Universal Robots URScript: Fuk_Rabbit_01D.script

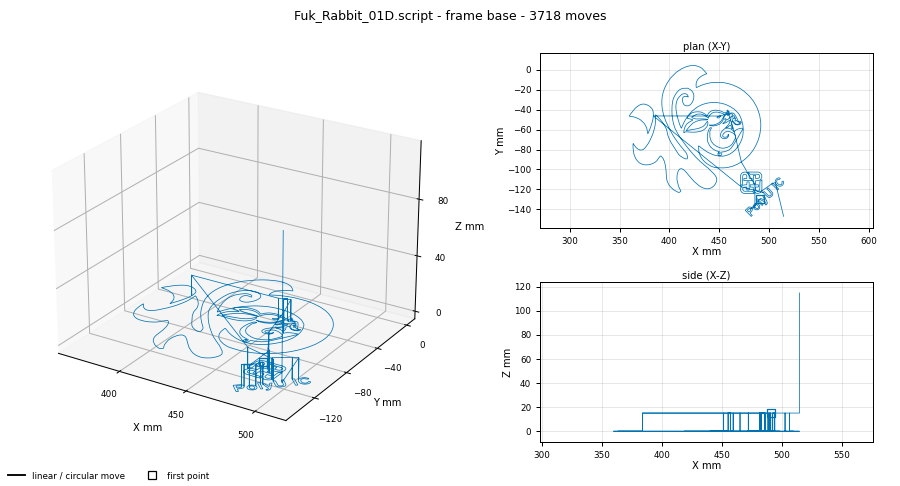
[picture p0: tool path of Fuk_Rabbit_01D.script in frame base, 3718 of 3719 moves have a stored position in this frame; points joined in program order, loops and branches not executed]
  global speed_ms    = 0.300
  global speed_rads  = 0.750
  global accel_mss   = 3.000
  global accel_radss = 1.200
  global blend_radius_m = 0.001




  # Main program:
  # Program generated by RoboDK v5.4.3 for UR10e on 11/01/2023 10:45:26
  # Using nominal kinematics.
  blend_radius_m = 0.001
  speed_ms    = 1.000
  # set_reference(p[0.514600, -0.147080, 0.000000, 0.000000, 0.000000, 1.570796])
  set_tcp(p[0.002800, -0.002800, 0.20500, 0.000000, 0.000000, 0.000000])
  movej([0.091562, -1.751682, -1.942220, -4.160080, -1.570796, -1.479235],accel_radss,speed_rads,0,0)
  movel(p[0.490670, -0.129830, 0.015000, 0.000000, -3.141593, 0.000000],accel_mss,speed_ms,0,0)

  speed_ms    = 1.000
  movel(p[0.490670, -0.129830, 0.015000, 0.000000, -3.141593, 0.000000],accel_mss,speed_ms,0,0.000)

  movel(p[0.490670, -0.129830, 0.003000, 0.000000, -3.141593, 0.000000],accel_mss,speed_ms,0,blend_radius_m)
  speed_ms    = 0.050
  movel(p[0.490670, -0.129830, -0.000100, 0.000000, -3.141593, 0.000000],accel_mss,speed_ms,0,blend_radius_m)
  speed_ms    = 0.083
  movel(p[0.491032, -0.129476, -0.000100, 0.000000, -3.141593, 0.000000],accel_mss,speed_ms,0,0.000)
  movel(p[0.491414, -0.129146, -0.000100, 0.000000, -3.141593, 0.000000],accel_mss,speed_ms,0,0.000)
  movel(p[0.491603, -0.129079, -0.000100, 0.000000, -3.141593, 0.000000],accel_mss,speed_ms,0,0.000)
  movel(p[0.491737, -0.129108, -0.000100, 0.000000, -3.141593, 0.000000],accel_mss,speed_ms,0,0.000)
  movel(p[0.492253, -0.129343, -0.000100, 0.000000, -3.141593, 0.000000],accel_mss,speed_ms,0,0.000)
  movel(p[0.492858, -0.129634, -0.000100, 0.000000, -3.141593, 0.000000],accel_mss,speed_ms,0,0.000)
  movel(p[0.493538, -0.129979, -0.000100, 0.000000, -3.141593, 0.000000],accel_mss,speed_ms,0,0.000)
  movel(p[0.494662, -0.130547, -0.000100, 0.000000, -3.141593, 0.000000],accel_mss,speed_ms,0,0.001)
  movel(p[0.495264, -0.130798, -0.000100, 0.000000, -3.141593, 0.000000],accel_mss,speed_ms,0,0.000)
  movel(p[0.495582, -0.130848, -0.000100, 0.000000, -3.141593, 0.000000],accel_mss,speed_ms,0,0.000)
  movel(p[0.495701, -0.130727, -0.000100, 0.000000, -3.141593, 0.000000],accel_mss,speed_ms,0,0.000)
  movel(p[0.495677, -0.130619, -0.000100, 0.000000, -3.141593, 0.000000],accel_mss,speed_ms,0,0.000)
  movel(p[0.495417, -0.130053, -0.000100, 0.000000, -3.141593, 0.000000],accel_mss,speed_ms,0,0.000)
  movel(p[0.495105, -0.129397, -0.000100, 0.000000, -3.141593, 0.000000],accel_mss,speed_ms,0,0.000)
  movel(p[0.494735, -0.128647, -0.000100, 0.000000, -3.141593, 0.000000],accel_mss,speed_ms,0,0.000)
  movel(p[0.494252, -0.127684, -0.000100, 0.000000, -3.141593, 0.000000],accel_mss,speed_ms,0,0.000)
  movel(p[0.493769, -0.126720, -0.000100, 0.000000, -3.141593, 0.000000],accel_mss,speed_ms,0,0.000)
  movel(p[0.494025, -0.126472, -0.000100, 0.000000, -3.141593, 0.000000],accel_mss,speed_ms,0,0.000)
  movel(p[0.494281, -0.126224, -0.000100, 0.000000, -3.141593, 0.000000],accel_mss,speed_ms,0,0.000)
  movel(p[0.494536, -0.125976, -0.000100, 0.000000, -3.141593, 0.000000],accel_mss,speed_ms,0,0.000)
  movel(p[0.494792, -0.125728, -0.000100, 0.000000, -3.141593, 0.000000],accel_mss,speed_ms,0,0.000)
  movel(p[0.495325, -0.126847, -0.000100, 0.000000, -3.141593, 0.000000],accel_mss,speed_ms,0,0.000)
  movel(p[0.495859, -0.127966, -0.000100, 0.000000, -3.141593, 0.000000],accel_mss,speed_ms,0,0.000)
  movel(p[0.496321, -0.128940, -0.000100, 0.000000, -3.141593, 0.000000],accel_mss,speed_ms,0,0.000)
  movel(p[0.496781, -0.129915, -0.000100, 0.000000, -3.141593, 0.000000],accel_mss,speed_ms,0,0.000)
  movel(p[0.497237, -0.130892, -0.000100, 0.000000, -3.141593, 0.000000],accel_mss,speed_ms,0,0.000)
  movel(p[0.497690, -0.131870, -0.000100, 0.000000, -3.141593, 0.000000],accel_mss,speed_ms,0,0.000)
  movel(p[0.498208, -0.133320, -0.000100, 0.000000, -3.141593, 0.000000],accel_mss,speed_ms,0,0.001)
  movel(p[0.498190, -0.134226, -0.000100, 0.000000, -3.141593, 0.000000],accel_mss,speed_ms,0,0.000)
  movel(p[0.497708, -0.135078, -0.000100, 0.000000, -3.141593, 0.000000],accel_mss,speed_ms,0,0.000)
  movel(p[0.497304, -0.135478, -0.000100, 0.000000, -3.141593, 0.000000],accel_mss,speed_ms,0,0.000)
  movel(p[0.497002, -0.135642, -0.000100, 0.000000, -3.141593, 0.000000],accel_mss,speed_ms,0,0.000)
  movel(p[0.496727, -0.135624, -0.000100, 0.000000, -3.141593, 0.000000],accel_mss,speed_ms,0,0.000)
  movel(p[0.496428, -0.135434, -0.000100, 0.000000, -3.141593, 0.000000],accel_mss,speed_ms,0,0.000)
  movel(p[0.496280, -0.135274, -0.000100, 0.000000, -3.141593, 0.000000],accel_mss,speed_ms,0,0.000)
  movel(p[0.496250, -0.135159, -0.000100, 0.000000, -3.141593, 0.000000],accel_mss,speed_ms,0,0.000)
  movel(p[0.496310, -0.135021, -0.000100, 0.000000, -3.141593, 0.000000],accel_mss,speed_ms,0,0.000)
  movel(p[0.496545, -0.134729, -0.000100, 0.000000, -3.141593, 0.000000],accel_mss,speed_ms,0,0.000)
  movel(p[0.496741, -0.134465, -0.000100, 0.000000, -3.141593, 0.000000],accel_mss,speed_ms,0,0.000)
  movel(p[0.496842, -0.134244, -0.000100, 0.000000, -3.141593, 0.000000],accel_mss,speed_ms,0,0.000)
  movel(p[0.496876, -0.134003, -0.000100, 0.000000, -3.141593, 0.000000],accel_mss,speed_ms,0,0.000)
  movel(p[0.496853, -0.133678, -0.000100, 0.000000, -3.141593, 0.000000],accel_mss,speed_ms,0,0.000)
  movel(p[0.496808, -0.133438, -0.000100, 0.000000, -3.141593, 0.000000],accel_mss,speed_ms,0,0.000)
  movel(p[0.496738, -0.133207, -0.000100, 0.000000, -3.141593, 0.000000],accel_mss,speed_ms,0,0.000)
  movel(p[0.496657, -0.133013, -0.000100, 0.000000, -3.141593, 0.000000],accel_mss,speed_ms,0,0.000)
  movel(p[0.496575, -0.132902, -0.000100, 0.000000, -3.141593, 0.000000],accel_mss,speed_ms,0,0.000)
  movel(p[0.496413, -0.132791, -0.000100, 0.000000, -3.141593, 0.000000],accel_mss,speed_ms,0,0.000)
  movel(p[0.495586, -0.132385, -0.000100, 0.000000, -3.141593, 0.000000],accel_mss,speed_ms,0,0.000)
  movel(p[0.494609, -0.131919, -0.000100, 0.000000, -3.141593, 0.000000],accel_mss,speed_ms,0,0.000)
  movel(p[0.493488, -0.131401, -0.000100, 0.000000, -3.141593, 0.000000],accel_mss,speed_ms,0,0.000)
  movel(p[0.492381, -0.130891, -0.000100, 0.000000, -3.141593, 0.000000],accel_mss,speed_ms,0,0.000)
  movel(p[0.491449, -0.130448, -0.000100, 0.000000, -3.141593, 0.000000],accel_mss,speed_ms,0,0.000)
  movel(p[0.490630, -0.130050, -0.000100, 0.000000, -3.141593, 0.000000],accel_mss,speed_ms,0,0.000)
  movel(p[0.490670, -0.129830, -0.000100, 0.000000, -3.141593, 0.000000],accel_mss,speed_ms,0,0.000)
  speed_ms    = 0.050
  movel(p[0.490670, -0.129830, 0.003000, 0.000000, -3.141593, 0.000000],accel_mss,speed_ms,0,blend_radius_m)
  speed_ms    = 1.000
  movel(p[0.490670, -0.129830, 0.015000, 0.000000, -3.141593, 0.000000],accel_mss,speed_ms,0,blend_radius_m)

  movel(p[0.489450, -0.130704, 0.015000, 0.000000, -3.141593, 0.000000],accel_mss,speed_ms,0,0.001)

  movel(p[0.489450, -0.130704, 0.003000, 0.000000, -3.141593, 0.000000],accel_mss,speed_ms,0,blend_radius_m)
  speed_ms    = 0.050
  movel(p[0.489450, -0.130704, -0.000100, 0.000000, -3.141593, 0.000000],accel_mss,speed_ms,0,blend_radius_m)
  speed_ms    = 0.083
  movel(p[0.490933, -0.132187, -0.000100, 0.000000, -3.141593, 0.000000],accel_mss,speed_ms,0,0.001)
  movel(p[0.492071, -0.133333, -0.000100, 0.000000, -3.141593, 0.000000],accel_mss,speed_ms,0,0.001)
  movel(p[0.493029, -0.134322, -0.000100, 0.000000, -3.141593, 0.000000],accel_mss,speed_ms,0,0.001)
  movel(p[0.493862, -0.135197, -0.000100, 0.000000, -3.141593, 0.000000],accel_mss,speed_ms,0,0.000)
  movel(p[0.493901, -0.135293, -0.000100, 0.000000, -3.141593, 0.000000],accel_mss,speed_ms,0,0.000)
  movel(p[0.493835, -0.135480, -0.000100, 0.000000, -3.141593, 0.000000],accel_mss,speed_ms,0,0.000)
  movel(p[0.493567, -0.135785, -0.000100, 0.000000, -3.141593, 0.000000],accel_mss,speed_ms,0,0.000)
  movel(p[0.493270, -0.136063, -0.000100, 0.000000, -3.141593, 0.000000],accel_mss,speed_ms,0,0.000)
  movel(p[0.493088, -0.136129, -0.000100, 0.000000, -3.141593, 0.000000],accel_mss,speed_ms,0,0.000)
  movel(p[0.492980, -0.136086, -0.000100, 0.000000, -3.141593, 0.000000],accel_mss,speed_ms,0,0.000)
  movel(p[0.492106, -0.135260, -0.000100, 0.000000, -3.141593, 0.000000],accel_mss,speed_ms,0,0.000)
  movel(p[0.491114, -0.134305, -0.000100, 0.000000, -3.141593, 0.000000],accel_mss,speed_ms,0,0.001)
  movel(p[0.489967, -0.133171, -0.000100, 0.000000, -3.141593, 0.000000],accel_mss,speed_ms,0,0.001)
  movel(p[0.488487, -0.131692, -0.000100, 0.000000, -3.141593, 0.000000],accel_mss,speed_ms,0,0.001)
  movel(p[0.487006, -0.130212, -0.000100, 0.000000, -3.141593, 0.000000],accel_mss,speed_ms,0,0.001)
  movel(p[0.487246, -0.129965, -0.000100, 0.000000, -3.141593, 0.000000],accel_mss,speed_ms,0,0.000)
  movel(p[0.487486, -0.129717, -0.000100, 0.000000, -3.141593, 0.000000],accel_mss,speed_ms,0,0.000)
  movel(p[0.487726, -0.129470, -0.000100, 0.000000, -3.141593, 0.000000],accel_mss,speed_ms,0,0.000)
  movel(p[0.487966, -0.129222, -0.000100, 0.000000, -3.141593, 0.000000],accel_mss,speed_ms,0,0.000)
  movel(p[0.489450, -0.130704, -0.000100, 0.000000, -3.141593, 0.000000],accel_mss,speed_ms,0,0.001)
  speed_ms    = 0.050
  movel(p[0.489450, -0.130704, 0.003000, 0.000000, -3.141593, 0.000000],accel_mss,speed_ms,0,blend_radius_m)
  speed_ms    = 1.000
  movel(p[0.489450, -0.130704, 0.015000, 0.000000, -3.141593, 0.000000],accel_mss,speed_ms,0,blend_radius_m)

  movel(p[0.488402, -0.134348, 0.015000, 0.000000, -3.141593, 0.000000],accel_mss,speed_ms,0,blend_radius_m)

  movel(p[0.488402, -0.134348, 0.003000, 0.000000, -3.141593, 0.000000],accel_mss,speed_ms,0,blend_radius_m)
  speed_ms    = 0.050
  movel(p[0.488402, -0.134348, -0.000100, 0.000000, -3.141593, 0.000000],accel_mss,speed_ms,0,blend_radius_m)
  speed_ms    = 0.083
  movel(p[0.489131, -0.134715, -0.000100, 0.000000, -3.141593, 0.000000],accel_mss,speed_ms,0,0.000)
  movel(p[0.489694, -0.135212, -0.000100, 0.000000, -3.141593, 0.000000],accel_mss,speed_ms,0,0.000)
  movel(p[0.490184, -0.135859, -0.000100, 0.000000, -3.141593, 0.000000],accel_mss,speed_ms,0,0.000)
  movel(p[0.490543, -0.136563, -0.000100, 0.000000, -3.141593, 0.000000],accel_mss,speed_ms,0,0.000)
  movel(p[0.490711, -0.137230, -0.000100, 0.000000, -3.141593, 0.000000],accel_mss,speed_ms,0,0.000)
  movel(p[0.490469, -0.138750, -0.000100, 0.000000, -3.141593, 0.000000],accel_mss,speed_ms,0,0.001)
  movel(p[0.489477, -0.139984, -0.000100, 0.000000, -3.141593, 0.000000],accel_mss,speed_ms,0,0.001)
  movel(p[0.488016, -0.140593, -0.000100, 0.000000, -3.141593, 0.000000],accel_mss,speed_ms,0,0.001)
  movel(p[0.486490, -0.140400, -0.000100, 0.000000, -3.141593, 0.000000],accel_mss,speed_ms,0,0.001)
  movel(p[0.485962, -0.140097, -0.000100, 0.000000, -3.141593, 0.000000],accel_mss,speed_ms,0,0.000)
  movel(p[0.485374, -0.139591, -0.000100, 0.000000, -3.141593, 0.000000],accel_mss,speed_ms,0,0.000)
  movel(p[0.484851, -0.139015, -0.000100, 0.000000, -3.141593, 0.000000],accel_mss,speed_ms,0,0.000)
  movel(p[0.484531, -0.138492, -0.000100, 0.000000, -3.141593, 0.000000],accel_mss,speed_ms,0,0.000)
  movel(p[0.484440, -0.138227, -0.000100, 0.000000, -3.141593, 0.000000],accel_mss,speed_ms,0,0.000)
  movel(p[0.484378, -0.137886, -0.000100, 0.000000, -3.141593, 0.000000],accel_mss,speed_ms,0,0.000)
  movel(p[0.484347, -0.137493, -0.000100, 0.000000, -3.141593, 0.000000],accel_mss,speed_ms,0,0.000)
  movel(p[0.484349, -0.137070, -0.000100, 0.000000, -3.141593, 0.000000],accel_mss,speed_ms,0,0.000)
  movel(p[0.484479, -0.136262, -0.000100, 0.000000, -3.141593, 0.000000],accel_mss,speed_ms,0,0.000)
  movel(p[0.484789, -0.135564, -0.000100, 0.000000, -3.141593, 0.000000],accel_mss,speed_ms,0,0.000)
  movel(p[0.485282, -0.134982, -0.000100, 0.000000, -3.141593, 0.000000],accel_mss,speed_ms,0,0.000)
  movel(p[0.485951, -0.134516, -0.000100, 0.000000, -3.141593, 0.000000],accel_mss,speed_ms,0,0.000)
  movel(p[0.486717, -0.134242, -0.000100, 0.000000, -3.141593, 0.000000],accel_mss,speed_ms,0,0.000)
  movel(p[0.487565, -0.134186, -0.000100, 0.000000, -3.141593, 0.000000],accel_mss,speed_ms,0,0.000)
  movel(p[0.488402, -0.134348, -0.000100, 0.000000, -3.141593, 0.000000],accel_mss,speed_ms,0,0.000)
  speed_ms    = 0.050
  movel(p[0.488402, -0.134348, 0.003000, 0.000000, -3.141593, 0.000000],accel_mss,speed_ms,0,blend_radius_m)
  speed_ms    = 1.000
  movel(p[0.488402, -0.134348, 0.015000, 0.000000, -3.141593, 0.000000],accel_mss,speed_ms,0,blend_radius_m)

  movel(p[0.482360, -0.138384, 0.015000, 0.000000, -3.141593, 0.000000],accel_mss,speed_ms,0,blend_radius_m)

  movel(p[0.482360, -0.138384, 0.003000, 0.000000, -3.141593, 0.000000],accel_mss,speed_ms,0,blend_radius_m)
  speed_ms    = 0.050
  movel(p[0.482360, -0.138384, -0.000100, 0.000000, -3.141593, 0.000000],accel_mss,speed_ms,0,blend_radius_m)
  speed_ms    = 0.083
  movel(p[0.482929, -0.139159, -0.000100, 0.000000, -3.141593, 0.000000],accel_mss,speed_ms,0,0.000)
  movel(p[0.483207, -0.140028, -0.000100, 0.000000, -3.141593, 0.000000],accel_mss,speed_ms,0,0.000)
  movel(p[0.483162, -0.140801, -0.000100, 0.000000, -3.141593, 0.000000],accel_mss,speed_ms,0,0.000)
  movel(p[0.482760, -0.141616, -0.000100, 0.000000, -3.141593, 0.000000],accel_mss,speed_ms,0,0.000)
  movel(p[0.481912, -0.142642, -0.000100, 0.000000, -3.141593, 0.000000],accel_mss,speed_ms,0,0.001)
  movel(p[0.481563, -0.143031, -0.000100, 0.000000, -3.141593, 0.000000],accel_mss,speed_ms,0,0.000)
  movel(p[0.481268, -0.143389, -0.000100, 0.000000, -3.141593, 0.000000],accel_mss,speed_ms,0,0.000)
  movel(p[0.481038, -0.143695, -0.000100, 0.000000, -3.141593, 0.000000],accel_mss,speed_ms,0,0.000)
  movel(p[0.481001, -0.143809, -0.000100, 0.000000, -3.141593, 0.000000],accel_mss,speed_ms,0,0.000)
  movel(p[0.481041, -0.143924, -0.000100, 0.000000, -3.141593, 0.000000],accel_mss,speed_ms,0,0.000)
  movel(p[0.481318, -0.144261, -0.000100, 0.000000, -3.141593, 0.000000],accel_mss,speed_ms,0,0.000)
  movel(p[0.481667, -0.144654, -0.000100, 0.000000, -3.141593, 0.000000],accel_mss,speed_ms,0,0.000)
  movel(p[0.482081, -0.145085, -0.000100, 0.000000, -3.141593, 0.000000],accel_mss,speed_ms,0,0.000)
  movel(p[0.482622, -0.145629, -0.000100, 0.000000, -3.141593, 0.000000],accel_mss,speed_ms,0,0.000)
  movel(p[0.483162, -0.146173, -0.000100, 0.000000, -3.141593, 0.000000],accel_mss,speed_ms,0,0.000)
  movel(p[0.482945, -0.146400, -0.000100, 0.000000, -3.141593, 0.000000],accel_mss,speed_ms,0,0.000)
  movel(p[0.482728, -0.146626, -0.000100, 0.000000, -3.141593, 0.000000],accel_mss,speed_ms,0,0.000)
  movel(p[0.482551, -0.146800, -0.000100, 0.000000, -3.141593, 0.000000],accel_mss,speed_ms,0,0.000)
  movel(p[0.482375, -0.146946, -0.000100, 0.000000, -3.141593, 0.000000],accel_mss,speed_ms,0,0.000)
  movel(p[0.482222, -0.147054, -0.000100, 0.000000, -3.141593, 0.000000],accel_mss,speed_ms,0,0.000)
  movel(p[0.482028, -0.147038, -0.000100, 0.000000, -3.141593, 0.000000],accel_mss,speed_ms,0,0.000)
  movel(p[0.481182, -0.146232, -0.000100, 0.000000, -3.141593, 0.000000],accel_mss,speed_ms,0,0.000)
  movel(p[0.480223, -0.145300, -0.000100, 0.000000, -3.141593, 0.000000],accel_mss,speed_ms,0,0.001)
  movel(p[0.479114, -0.144192, -0.000100, 0.000000, -3.141593, 0.000000],accel_mss,speed_ms,0,0.001)
  movel(p[0.478015, -0.143074, -0.000100, 0.000000, -3.141593, 0.000000],accel_mss,speed_ms,0,0.001)
  movel(p[0.477085, -0.142106, -0.000100, 0.000000, -3.141593, 0.000000],accel_mss,speed_ms,0,0.001)
  movel(p[0.476280, -0.141253, -0.000100, 0.000000, -3.141593, 0.000000],accel_mss,speed_ms,0,0.000)
  movel(p[0.476227, -0.141145, -0.000100, 0.000000, -3.141593, 0.000000],accel_mss,speed_ms,0,0.000)
  movel(p[0.476318, -0.140864, -0.000100, 0.000000, -3.141593, 0.000000],accel_mss,speed_ms,0,0.000)
  movel(p[0.477774, -0.139443, -0.000100, 0.000000, -3.141593, 0.000000],accel_mss,speed_ms,0,0.001)
  movel(p[0.479184, -0.138110, -0.000100, 0.000000, -3.141593, 0.000000],accel_mss,speed_ms,0,0.001)
  movel(p[0.479706, -0.137786, -0.000100, 0.000000, -3.141593, 0.000000],accel_mss,speed_ms,0,0.000)
  movel(p[0.480611, -0.137640, -0.000100, 0.000000, -3.141593, 0.000000],accel_mss,speed_ms,0,0.000)
  movel(p[0.481544, -0.137852, -0.000100, 0.000000, -3.141593, 0.000000],accel_mss,speed_ms,0,0.000)
  movel(p[0.482360, -0.138384, -0.000100, 0.000000, -3.141593, 0.000000],accel_mss,speed_ms,0,0.000)
  speed_ms    = 0.050
  movel(p[0.482360, -0.138384, 0.003000, 0.000000, -3.141593, 0.000000],accel_mss,speed_ms,0,blend_radius_m)
  speed_ms    = 1.000
  movel(p[0.482360, -0.138384, 0.015000, 0.000000, -3.141593, 0.000000],accel_mss,speed_ms,0,blend_radius_m)

  movel(p[0.481296, -0.139556, 0.015000, 0.000000, -3.141593, 0.000000],accel_mss,speed_ms,0,0.001)

  movel(p[0.481296, -0.139556, 0.003000, 0.000000, -3.141593, 0.000000],accel_mss,speed_ms,0,blend_radius_m)
  speed_ms    = 0.050
  movel(p[0.481296, -0.139556, -0.000100, 0.000000, -3.141593, 0.000000],accel_mss,speed_ms,0,blend_radius_m)
  speed_ms    = 0.083
  movel(p[0.481636, -0.140114, -0.000100, 0.000000, -3.141593, 0.000000],accel_mss,speed_ms,0,0.000)
  movel(p[0.481657, -0.140724, -0.000100, 0.000000, -3.141593, 0.000000],accel_mss,speed_ms,0,0.000)
  movel(p[0.481568, -0.140933, -0.000100, 0.000000, -3.141593, 0.000000],accel_mss,speed_ms,0,0.000)
  movel(p[0.481354, -0.141251, -0.000100, 0.000000, -3.141593, 0.000000],accel_mss,speed_ms,0,0.000)
  movel(p[0.481077, -0.141604, -0.000100, 0.000000, -3.141593, 0.000000],accel_mss,speed_ms,0,0.000)
  movel(p[0.480768, -0.141945, -0.000100, 0.000000, -3.141593, 0.000000],accel_mss,speed_ms,0,0.000)
  movel(p[0.480163, -0.142512, -0.000100, 0.000000, -3.141593, 0.000000],accel_mss,speed_ms,0,0.000)
  movel(p[0.479815, -0.142622, -0.000100, 0.000000, -3.141593, 0.000000],accel_mss,speed_ms,0,0.000)
  movel(p[0.479457, -0.142458, -0.000100, 0.000000, -3.141593, 0.000000],accel_mss,speed_ms,0,0.000)
  movel(p[0.478765, -0.141753, -0.000100, 0.000000, -3.141593, 0.000000],accel_mss,speed_ms,0,0.000)
  movel(p[0.478330, -0.141231, -0.000100, 0.000000, -3.141593, 0.000000],accel_mss,speed_ms,0,0.000)
  movel(p[0.478275, -0.140954, -0.000100, 0.000000, -3.141593, 0.000000],accel_mss,speed_ms,0,0.000)
  movel(p[0.478446, -0.140660, -0.000100, 0.000000, -3.141593, 0.000000],accel_mss,speed_ms,0,0.000)
  movel(p[0.479256, -0.139890, -0.000100, 0.000000, -3.141593, 0.000000],accel_mss,speed_ms,0,0.000)
  movel(p[0.479504, -0.139676, -0.000100, 0.000000, -3.141593, 0.000000],accel_mss,speed_ms,0,0.000)
  movel(p[0.479770, -0.139475, -0.000100, 0.000000, -3.141593, 0.000000],accel_mss,speed_ms,0,0.000)
  movel(p[0.480015, -0.139313, -0.000100, 0.000000, -3.141593, 0.000000],accel_mss,speed_ms,0,0.000)
  movel(p[0.480188, -0.139231, -0.000100, 0.000000, -3.141593, 0.000000],accel_mss,speed_ms,0,0.000)
  movel(p[0.480757, -0.139223, -0.000100, 0.000000, -3.141593, 0.000000],accel_mss,speed_ms,0,0.000)
  movel(p[0.481296, -0.139556, -0.000100, 0.000000, -3.141593, 0.000000],accel_mss,speed_ms,0,0.000)
  speed_ms    = 0.050
  movel(p[0.481296, -0.139556, 0.003000, 0.000000, -3.141593, 0.000000],accel_mss,speed_ms,0,blend_radius_m)
  speed_ms    = 1.000
  movel(p[0.481296, -0.139556, 0.015000, 0.000000, -3.141593, 0.000000],accel_mss,speed_ms,0,blend_radius_m)

  movel(p[0.485804, -0.137802, 0.015000, 0.000000, -3.141593, 0.000000],accel_mss,speed_ms,0,blend_radius_m)

  movel(p[0.485804, -0.137802, 0.003000, 0.000000, -3.141593, 0.000000],accel_mss,speed_ms,0,blend_radius_m)
  speed_ms    = 0.050
  movel(p[0.485804, -0.137802, -0.000100, 0.000000, -3.141593, 0.000000],accel_mss,speed_ms,0,blend_radius_m)
  speed_ms    = 0.083
  movel(p[0.485574, -0.137101, -0.000100, 0.000000, -3.141593, 0.000000],accel_mss,speed_ms,0,0.000)
  movel(p[0.485633, -0.136451, -0.000100, 0.000000, -3.141593, 0.000000],accel_mss,speed_ms,0,0.000)
  movel(p[0.485964, -0.135890, -0.000100, 0.000000, -3.141593, 0.000000],accel_mss,speed_ms,0,0.000)
  movel(p[0.486573, -0.135499, -0.000100, 0.000000, -3.141593, 0.000000],accel_mss,speed_ms,0,0.000)
  movel(p[0.487296, -0.135441, -0.000100, 0.000000, -3.141593, 0.000000],accel_mss,speed_ms,0,0.000)
  movel(p[0.488060, -0.135741, -0.000100, 0.000000, -3.141593, 0.000000],accel_mss,speed_ms,0,0.000)
  movel(p[0.488778, -0.136364, -0.000100, 0.000000, -3.141593, 0.000000],accel_mss,speed_ms,0,0.000)
  movel(p[0.489185, -0.136902, -0.000100, 0.000000, -3.141593, 0.000000],accel_mss,speed_ms,0,0.000)
  movel(p[0.489414, -0.137395, -0.000100, 0.000000, -3.141593, 0.000000],accel_mss,speed_ms,0,0.000)
  movel(p[0.489476, -0.137873, -0.000100, 0.000000, -3.141593, 0.000000],accel_mss,speed_ms,0,0.000)
  movel(p[0.489384, -0.138362, -0.000100, 0.000000, -3.141593, 0.000000],accel_mss,speed_ms,0,0.000)
  movel(p[0.488887, -0.139008, -0.000100, 0.000000, -3.141593, 0.000000],accel_mss,speed_ms,0,0.000)
  movel(p[0.488066, -0.139280, -0.000100, 0.000000, -3.141593, 0.000000],accel_mss,speed_ms,0,0.000)
  movel(p[0.487122, -0.139099, -0.000100, 0.000000, -3.141593, 0.000000],accel_mss,speed_ms,0,0.000)
  movel(p[0.486306, -0.138506, -0.000100, 0.000000, -3.141593, 0.000000],accel_mss,speed_ms,0,0.000)
  movel(p[0.485804, -0.137802, -0.000100, 0.000000, -3.141593, 0.000000],accel_mss,speed_ms,0,0.000)
  speed_ms    = 0.050
  movel(p[0.485804, -0.137802, 0.003000, 0.000000, -3.141593, 0.000000],accel_mss,speed_ms,0,blend_radius_m)
  speed_ms    = 1.000
  movel(p[0.485804, -0.137802, 0.015000, 0.000000, -3.141593, 0.000000],accel_mss,speed_ms,0,blend_radius_m)

  movel(p[0.485801, -0.114304, 0.015000, 0.000000, -3.141593, 0.000000],accel_mss,speed_ms,0,blend_radius_m)

  movel(p[0.485801, -0.114304, 0.003000, 0.000000, -3.141593, 0.000000],accel_mss,speed_ms,0,blend_radius_m)
  speed_ms    = 0.050
  movel(p[0.485801, -0.114304, -0.000100, 0.000000, -3.141593, 0.000000],accel_mss,speed_ms,0,blend_radius_m)
  speed_ms    = 0.083
  movel(p[0.485276, -0.114304, -0.000100, 0.000000, -3.141593, 0.000000],accel_mss,speed_ms,0,0.000)
  movel(p[0.484751, -0.114304, -0.000100, 0.000000, -3.141593, 0.000000],accel_mss,speed_ms,0,0.000)
  movel(p[0.484226, -0.114304, -0.000100, 0.000000, -3.141593, 0.000000],accel_mss,speed_ms,0,0.000)
  movel(p[0.484226, -0.112241, -0.000100, 0.000000, -3.141593, 0.000000],accel_mss,speed_ms,0,0.001)
  movel(p[0.484226, -0.110179, -0.000100, 0.000000, -3.141593, 0.000000],accel_mss,speed_ms,0,0.001)
  movel(p[0.484226, -0.108116, -0.000100, 0.000000, -3.141593, 0.000000],accel_mss,speed_ms,0,0.001)
  movel(p[0.484226, -0.106054, -0.000100, 0.000000, -3.141593, 0.000000],accel_mss,speed_ms,0,0.001)
  movel(p[0.484769, -0.106032, -0.000100, 0.000000, -3.141593, 0.000000],accel_mss,speed_ms,0,0.000)
  movel(p[0.485313, -0.106010, -0.000100, 0.000000, -3.141593, 0.000000],accel_mss,speed_ms,0,0.000)
  movel(p[0.485857, -0.105988, -0.000100, 0.000000, -3.141593, 0.000000],accel_mss,speed_ms,0,0.000)
  movel(p[0.486401, -0.105966, -0.000100, 0.000000, -3.141593, 0.000000],accel_mss,speed_ms,0,0.000)
  movel(p[0.486401, -0.106719, -0.000100, 0.000000, -3.141593, 0.000000],accel_mss,speed_ms,0,0.000)
  movel(p[0.486401, -0.107472, -0.000100, 0.000000, -3.141593, 0.000000],accel_mss,speed_ms,0,0.000)
  movel(p[0.486401, -0.108226, -0.000100, 0.000000, -3.141593, 0.000000],accel_mss,speed_ms,0,0.000)
  movel(p[0.486401, -0.108979, -0.000100, 0.000000, -3.141593, 0.000000],accel_mss,speed_ms,0,0.000)
  movel(p[0.487094, -0.108979, -0.000100, 0.000000, -3.141593, 0.000000],accel_mss,speed_ms,0,0.000)
  movel(p[0.487788, -0.108978, -0.000100, 0.000000, -3.141593, 0.000000],accel_mss,speed_ms,0,0.000)
  movel(p[0.488520, -0.108965, -0.000100, 0.000000, -3.141593, 0.000000],accel_mss,speed_ms,0,0.000)
  movel(p[0.488995, -0.108919, -0.000100, 0.000000, -3.141593, 0.000000],accel_mss,speed_ms,0,0.000)
  movel(p[0.489346, -0.108831, -0.000100, 0.000000, -3.141593, 0.000000],accel_mss,speed_ms,0,0.000)
  movel(p[0.489656, -0.108685, -0.000100, 0.000000, -3.141593, 0.000000],accel_mss,speed_ms,0,0.000)
  movel(p[0.490385, -0.107906, -0.000100, 0.000000, -3.141593, 0.000000],accel_mss,speed_ms,0,0.000)
  movel(p[0.490630, -0.106843, -0.000100, 0.000000, -3.141593, 0.000000],accel_mss,speed_ms,0,0.000)
  movel(p[0.490325, -0.105795, -0.000100, 0.000000, -3.141593, 0.000000],accel_mss,speed_ms,0,0.000)
  movel(p[0.489553, -0.105058, -0.000100, 0.000000, -3.141593, 0.000000],accel_mss,speed_ms,0,0.000)
  movel(p[0.489106, -0.104903, -0.000100, 0.000000, -3.141593, 0.000000],accel_mss,speed_ms,0,0.000)
  movel(p[0.488451, -0.104824, -0.000100, 0.000000, -3.141593, 0.000000],accel_mss,speed_ms,0,0.000)
  movel(p[0.487340, -0.104787, -0.000100, 0.000000, -3.141593, 0.000000],accel_mss,speed_ms,0,0.000)
  movel(p[0.484891, -0.104779, -0.000100, 0.000000, -3.141593, 0.000000],accel_mss,speed_ms,0,0.001)
  movel(p[0.482821, -0.104779, -0.000100, 0.000000, -3.141593, 0.000000],accel_mss,speed_ms,0,0.001)
  movel(p[0.480751, -0.104779, -0.000100, 0.000000, -3.141593, 0.000000],accel_mss,speed_ms,0,0.001)
  movel(p[0.480520, -0.104423, -0.000100, 0.000000, -3.141593, 0.000000],accel_mss,speed_ms,0,0.000)
  movel(p[0.480289, -0.104066, -0.000100, 0.000000, -3.141593, 0.000000],accel_mss,speed_ms,0,0.000)
  movel(p[0.480083, -0.103766, -0.000100, 0.000000, -3.141593, 0.000000],accel_mss,speed_ms,0,0.000)
  movel(p[0.479845, -0.103453, -0.000100, 0.000000, 3.141593, 0.000000],accel_mss,speed_ms,0,0.000)
  movel(p[0.479612, -0.103172, -0.000100, 0.000000, -3.141593, 0.000000],accel_mss,speed_ms,0,0.000)
  movel(p[0.479426, -0.102979, -0.000100, 0.000000, -3.141593, 0.000000],accel_mss,speed_ms,0,0.000)
  movel(p[0.479226, -0.102791, -0.000100, 0.000000, -3.141593, 0.000000],accel_mss,speed_ms,0,0.000)
  movel(p[0.479026, -0.102604, -0.000100, 0.000000, -3.141593, 0.000000],accel_mss,speed_ms,0,0.000)
  movel(p[0.481522, -0.102584, -0.000100, 0.000000, -3.141593, 0.000000],accel_mss,speed_ms,0,0.001)
  movel(p[0.484018, -0.102564, -0.000100, 0.000000, -3.141593, 0.000000],accel_mss,speed_ms,0,0.001)
  movel(p[0.486672, -0.102553, -0.000100, 0.000000, -3.141593, 0.000000],accel_mss,speed_ms,0,blend_radius_m)
  movel(p[0.488189, -0.102576, -0.000100, 0.000000, -3.141593, 0.000000],accel_mss,speed_ms,0,0.001)
  movel(p[0.489166, -0.102634, -0.000100, 0.000000, -3.141593, 0.000000],accel_mss,speed_ms,0,0.000)
  movel(p[0.489779, -0.102749, -0.000100, 0.000000, -3.141593, 0.000000],accel_mss,speed_ms,0,0.000)
  movel(p[0.491653, -0.103889, -0.000100, 0.000000, -3.141593, 0.000000],accel_mss,speed_ms,0,0.001)
  movel(p[0.492720, -0.105828, -0.000100, 0.000000, -3.141593, 0.000000],accel_mss,speed_ms,0,0.001)
  movel(p[0.492698, -0.108049, -0.000100, 0.000000, -3.141593, 0.000000],accel_mss,speed_ms,0,0.001)
  movel(p[0.491589, -0.109960, -0.000100, 0.000000, -3.141593, 0.000000],accel_mss,speed_ms,0,0.001)
  movel(p[0.490862, -0.110565, -0.000100, 0.000000, -3.141593, 0.000000],accel_mss,speed_ms,0,0.000)
  movel(p[0.490106, -0.110956, -0.000100, 0.000000, -3.141593, 0.000000],accel_mss,speed_ms,0,0.000)
  movel(p[0.489171, -0.111195, -0.000100, 0.000000, -3.141593, 0.000000],accel_mss,speed_ms,0,0.000)
  movel(p[0.487868, -0.111333, -0.000100, 0.000000, -3.141593, 0.000000],accel_mss,speed_ms,0,0.001)
  movel(p[0.487140, -0.111378, -0.000100, 0.000000, -3.141593, 0.000000],accel_mss,speed_ms,0,0.000)
  movel(p[0.486411, -0.111424, -0.000100, 0.000000, -3.141593, 0.000000],accel_mss,speed_ms,0,0.000)
  movel(p[0.486390, -0.112144, -0.000100, 0.000000, -3.141593, 0.000000],accel_mss,speed_ms,0,0.000)
  movel(p[0.486368, -0.112864, -0.000100, 0.000000, -3.141593, 0.000000],accel_mss,speed_ms,0,0.000)
  movel(p[0.486347, -0.113584, -0.000100, 0.000000, -3.141593, 0.000000],accel_mss,speed_ms,0,0.000)
  movel(p[0.486326, -0.114304, -0.000100, 0.000000, -3.141593, 0.000000],accel_mss,speed_ms,0,0.000)
  movel(p[0.485801, -0.114304, -0.000100, 0.000000, -3.141593, 0.000000],accel_mss,speed_ms,0,0.000)
  speed_ms    = 0.050
  movel(p[0.485801, -0.114304, 0.003000, 0.000000, -3.141593, 0.000000],accel_mss,speed_ms,0,blend_radius_m)
  speed_ms    = 1.000
  movel(p[0.485801, -0.114304, 0.015000, 0.000000, -3.141593, 0.000000],accel_mss,speed_ms,0,blend_radius_m)

  movel(p[0.483026, -0.111154, 0.015000, 0.000000, -3.141593, 0.000000],accel_mss,speed_ms,0,blend_radius_m)

  movel(p[0.483026, -0.111154, 0.003000, 0.000000, -3.141593, 0.000000],accel_mss,speed_ms,0,blend_radius_m)
  speed_ms    = 0.050
  movel(p[0.483026, -0.111154, -0.000100, 0.000000, -3.141593, 0.000000],accel_mss,speed_ms,0,blend_radius_m)
  speed_ms    = 0.083
  movel(p[0.480941, -0.111174, -0.000100, 0.000000, -3.141593, 0.000000],accel_mss,speed_ms,0,0.001)
  movel(p[0.478857, -0.111194, -0.000100, 0.000000, -3.141593, 0.000000],accel_mss,speed_ms,0,0.001)
  movel(p[0.476772, -0.111214, -0.000100, 0.000000, -3.141593, 0.000000],accel_mss,speed_ms,0,0.001)
  movel(p[0.474687, -0.111234, -0.000100, 0.000000, -3.141593, 0.000000],accel_mss,speed_ms,0,0.001)
  movel(p[0.474709, -0.110689, -0.000100, 0.000000, -3.141593, 0.000000],accel_mss,speed_ms,0,0.000)
  movel(p[0.474732, -0.110144, -0.000100, 0.000000, -3.141593, 0.000000],accel_mss,speed_ms,0,0.000)
  movel(p[0.474754, -0.109599, -0.000100, 0.000000, -3.141593, 0.000000],accel_mss,speed_ms,0,0.000)
  movel(p[0.474776, -0.109054, -0.000100, 0.000000, -3.141593, 0.000000],accel_mss,speed_ms,0,0.000)
  movel(p[0.475507, -0.109032, -0.000100, 0.000000, -3.141593, 0.000000],accel_mss,speed_ms,0,0.000)
  movel(p[0.476238, -0.109011, -0.000100, 0.000000, -3.141593, 0.000000],accel_mss,speed_ms,0,0.000)
  movel(p[0.476969, -0.108990, -0.000100, 0.000000, -3.141593, 0.000000],accel_mss,speed_ms,0,0.000)
  movel(p[0.477701, -0.108968, -0.000100, 0.000000, -3.141593, 0.000000],accel_mss,speed_ms,0,0.000)
  movel(p[0.477700, -0.108277, -0.000100, 0.000000, -3.141593, 0.000000],accel_mss,speed_ms,0,0.000)
  movel(p[0.477700, -0.107586, -0.000100, 0.000000, -3.141593, 0.000000],accel_mss,speed_ms,0,0.000)
  movel(p[0.477649, -0.106537, -0.000100, 0.000000, -3.141593, 0.000000],accel_mss,speed_ms,0,0.000)
  movel(p[0.477475, -0.105859, -0.000100, 0.000000, -3.141593, 0.000000],accel_mss,speed_ms,0,0.000)
  movel(p[0.477144, -0.105391, -0.000100, 0.000000, -3.141593, 0.000000],accel_mss,speed_ms,0,0.000)
  movel(p[0.476608, -0.105029, -0.000100, 0.000000, -3.141593, 0.000000],accel_mss,speed_ms,0,0.000)
  movel(p[0.475817, -0.104809, -0.000100, 0.000000, -3.141593, 0.000000],accel_mss,speed_ms,0,0.000)
  movel(p[0.475035, -0.104883, -0.000100, 0.000000, -3.141593, 0.000000],accel_mss,speed_ms,0,0.000)
  movel(p[0.474340, -0.105249, -0.000100, 0.000000, -3.141593, 0.000000],accel_mss,speed_ms,0,0.000)
  movel(p[0.473800, -0.105865, -0.000100, 0.000000, -3.141593, 0.000000],accel_mss,speed_ms,0,0.000)
  movel(p[0.473630, -0.106294, -0.000100, 0.000000, -3.141593, 0.000000],accel_mss,speed_ms,0,0.000)
  movel(p[0.473546, -0.106913, -0.000100, 0.000000, -3.141593, 0.000000],accel_mss,speed_ms,0,0.000)
  movel(p[0.473509, -0.107994, -0.000100, 0.000000, -3.141593, 0.000000],accel_mss,speed_ms,0,0.000)
  movel(p[0.473501, -0.110591, -0.000100, 0.000000, -3.141593, 0.000000],accel_mss,speed_ms,0,blend_radius_m)
  movel(p[0.473492, -0.112333, -0.000100, 0.000000, -3.141593, 0.000000],accel_mss,speed_ms,0,0.001)
  movel(p[0.473462, -0.113673, -0.000100, 0.000000, -3.141593, 0.000000],accel_mss,speed_ms,0,0.001)
  movel(p[0.473422, -0.114768, -0.000100, 0.000000, -3.141593, 0.000000],accel_mss,speed_ms,0,0.000)
  movel(p[0.473267, -0.114855, -0.000100, 0.000000, -3.141593, 0.000000],accel_mss,speed_ms,0,0.000)
  movel(p[0.472967, -0.115049, -0.000100, 0.000000, -3.141593, 0.000000],accel_mss,speed_ms,0,0.000)
  movel(p[0.472615, -0.115292, -0.000100, 0.000000, -3.141593, 0.000000],accel_mss,speed_ms,0,0.000)
  movel(p[0.472225, -0.115580, -0.000100, 0.000000, -3.141593, 0.000000],accel_mss,speed_ms,0,0.000)
  movel(p[0.471729, -0.115955, -0.000100, 0.000000, -3.141593, 0.000000],accel_mss,speed_ms,0,0.000)
  movel(p[0.471233, -0.116330, -0.000100, 0.000000, -3.141593, 0.000000],accel_mss,speed_ms,0,0.000)
  movel(p[0.471256, -0.113724, -0.000100, 0.000000, -3.141593, 0.000000],accel_mss,speed_ms,0,blend_radius_m)
  movel(p[0.471279, -0.111117, -0.000100, 0.000000, -3.141593, 0.000000],accel_mss,speed_ms,0,blend_radius_m)
  movel(p[0.471315, -0.107864, -0.000100, 0.000000, -3.141593, 0.000000],accel_mss,speed_ms,0,blend_radius_m)
  movel(p[0.471365, -0.106553, -0.000100, 0.000000, -3.141593, 0.000000],accel_mss,speed_ms,0,0.001)
  movel(p[0.471460, -0.105791, -0.000100, 0.000000, 3.141593, 0.000000],accel_mss,speed_ms,0,0.000)
  movel(p[0.471646, -0.105211, -0.000100, 0.000000, -3.141593, 0.000000],accel_mss,speed_ms,0,0.000)
  movel(p[0.472344, -0.104101, -0.000100, 0.000000, -3.141593, 0.000000],accel_mss,speed_ms,0,0.001)
  movel(p[0.473264, -0.103283, -0.000100, 0.000000, -3.141593, 0.000000],accel_mss,speed_ms,0,0.000)
  movel(p[0.474386, -0.102785, -0.000100, 0.000000, -3.141593, 0.000000],accel_mss,speed_ms,0,0.000)
  movel(p[0.475676, -0.102614, -0.000100, 0.000000, -3.141593, 0.000000],accel_mss,speed_ms,0,0.001)
  movel(p[0.476925, -0.102772, -0.000100, 0.000000, -3.141593, 0.000000],accel_mss,speed_ms,0,0.001)
  movel(p[0.478019, -0.103241, -0.000100, 0.000000, -3.141593, 0.000000],accel_mss,speed_ms,0,0.000)
  movel(p[0.478916, -0.104009, -0.000100, 0.000000, -3.141593, 0.000000],accel_mss,speed_ms,0,0.000)
  movel(p[0.479587, -0.105042, -0.000100, 0.000000, -3.141593, 0.000000],accel_mss,speed_ms,0,0.000)
  movel(p[0.479793, -0.105543, -0.000100, 0.000000, -3.141593, 0.000000],accel_mss,speed_ms,0,0.000)
  movel(p[0.479923, -0.106022, -0.000100, 0.000000, -3.141593, 0.000000],accel_mss,speed_ms,0,0.000)
  movel(p[0.480006, -0.106596, -0.000100, 0.000000, -3.141593, 0.000000],accel_mss,speed_ms,0,0.000)
  movel(p[0.480064, -0.107427, -0.000100, 0.000000, -3.141593, 0.000000],accel_mss,speed_ms,0,0.000)
  movel(p[0.480104, -0.108198, -0.000100, 0.000000, -3.141593, 0.000000],accel_mss,speed_ms,0,0.000)
  movel(p[0.480143, -0.108969, -0.000100, 0.000000, -3.141593, 0.000000],accel_mss,speed_ms,0,0.000)
  movel(p[0.480864, -0.108990, -0.000100, 0.000000, -3.141593, 0.000000],accel_mss,speed_ms,0,0.000)
  movel(p[0.481584, -0.109011, -0.000100, 0.000000, -3.141593, 0.000000],accel_mss,speed_ms,0,0.000)
  movel(p[0.482305, -0.109033, -0.000100, 0.000000, -3.141593, 0.000000],accel_mss,speed_ms,0,0.000)
  movel(p[0.483026, -0.109054, -0.000100, 0.000000, -3.141593, 0.000000],accel_mss,speed_ms,0,0.000)
  movel(p[0.483026, -0.109579, -0.000100, 0.000000, -3.141593, 0.000000],accel_mss,speed_ms,0,0.000)
  movel(p[0.483026, -0.110104, -0.000100, 0.000000, -3.141593, 0.000000],accel_mss,speed_ms,0,0.000)
  movel(p[0.483026, -0.110629, -0.000100, 0.000000, -3.141593, 0.000000],accel_mss,speed_ms,0,0.000)
  movel(p[0.483026, -0.111154, -0.000100, 0.000000, -3.141593, 0.000000],accel_mss,speed_ms,0,0.000)
  speed_ms    = 0.050
  movel(p[0.483026, -0.111154, 0.003000, 0.000000, -3.141593, 0.000000],accel_mss,speed_ms,0,blend_radius_m)
  speed_ms    = 1.000
  movel(p[0.483026, -0.111154, 0.015000, 0.000000, -3.141593, 0.000000],accel_mss,speed_ms,0,blend_radius_m)

  movel(p[0.472179, -0.092457, 0.015000, 0.000000, -3.141593, 0.000000],accel_mss,speed_ms,0,blend_radius_m)

  movel(p[0.472179, -0.092457, 0.003000, 0.000000, -3.141593, 0.000000],accel_mss,speed_ms,0,blend_radius_m)
  speed_ms    = 0.050
  movel(p[0.472179, -0.092457, -0.000100, 0.000000, -3.141593, 0.000000],accel_mss,speed_ms,0,blend_radius_m)
  speed_ms    = 0.083
  movel(p[0.472016, -0.092500, -0.000100, 0.000000, -3.141593, 0.000000],accel_mss,speed_ms,0,0.000)
  movel(p[0.471842, -0.092597, -0.000100, 0.000000, -3.141593, 0.000000],accel_mss,speed_ms,0,0.000)
  movel(p[0.471639, -0.092728, -0.000100, 0.000000, -3.141593, 0.000000],accel_mss,speed_ms,0,0.000)
  movel(p[0.471426, -0.092882, -0.000100, 0.000000, -3.141593, 0.000000],accel_mss,speed_ms,0,0.000)
  movel(p[0.471169, -0.093063, -0.000100, 0.000000, -3.141593, 0.000000],accel_mss,speed_ms,0,0.000)
  movel(p[0.470829, -0.093276, -0.000100, 0.000000, -3.141593, 0.000000],accel_mss,speed_ms,0,0.000)
  movel(p[0.470466, -0.093486, -0.000100, 0.000000, -3.141593, 0.000000],accel_mss,speed_ms,0,0.000)
  movel(p[0.470136, -0.093659, -0.000100, 0.000000, -3.141593, 0.000000],accel_mss,speed_ms,0,0.000)
  movel(p[0.469811, -0.093828, -0.000100, 0.000000, -3.141593, 0.000000],accel_mss,speed_ms,0,0.000)
  movel(p[0.469463, -0.094026, -0.000100, 0.000000, -3.141593, 0.000000],accel_mss,speed_ms,0,0.000)
  movel(p[0.469143, -0.094221, -0.000100, 0.000000, -3.141593, 0.000000],accel_mss,speed_ms,0,0.000)
  movel(p[0.468911, -0.094381, -0.000100, 0.000000, -3.141593, 0.000000],accel_mss,speed_ms,0,0.000)
  movel(p[0.468725, -0.094514, -0.000100, 0.000000, -3.141593, 0.000000],accel_mss,speed_ms,0,0.000)
  movel(p[0.468547, -0.094627, -0.000100, 0.000000, -3.141593, 0.000000],accel_mss,speed_ms,0,0.000)
  movel(p[0.468396, -0.094711, -0.000100, 0.000000, -3.141593, 0.000000],accel_mss,speed_ms,0,0.000)
  movel(p[0.468241, -0.094745, -0.000100, 0.000000, -3.141593, 0.000000],accel_mss,speed_ms,0,0.000)
  movel(p[0.467968, -0.094857, -0.000100, 0.000000, -3.141593, 0.000000],accel_mss,speed_ms,0,0.000)
  movel(p[0.467646, -0.094998, -0.000100, 0.000000, -3.141593, 0.000000],accel_mss,speed_ms,0,0.000)
  movel(p[0.467287, -0.095165, -0.000100, 0.000000, -3.141593, 0.000000],accel_mss,speed_ms,0,0.000)
  movel(p[0.465973, -0.095759, -0.000100, 0.000000, 3.141593, 0.000000],accel_mss,speed_ms,0,0.001)
  movel(p[0.464493, -0.096362, -0.000100, 0.000000, -3.141593, 0.000000],accel_mss,speed_ms,0,0.001)
  movel(p[0.463131, -0.096869, -0.000100, 0.000000, 3.141593, 0.000000],accel_mss,speed_ms,0,0.001)
  movel(p[0.462401, -0.097063, -0.000100, 0.000000, -3.141593, 0.000000],accel_mss,speed_ms,0,0.000)
  movel(p[0.462168, -0.097112, -0.000100, 0.000000, -3.141593, 0.000000],accel_mss,speed_ms,0,0.000)
  movel(p[0.461629, -0.097243, -0.000100, 0.000000, -3.141593, 0.000000],accel_mss,speed_ms,0,0.000)
  movel(p[0.460989, -0.097403, -0.000100, 0.000000, -3.141593, 0.000000],accel_mss,speed_ms,0,0.000)
  movel(p[0.460301, -0.097581, -0.000100, 0.000000, -3.141593, 0.000000],accel_mss,speed_ms,0,0.000)
  movel(p[0.458244, -0.098017, -0.000100, 0.000000, -3.141593, 0.000000],accel_mss,speed_ms,0,0.001)
  movel(p[0.455998, -0.098299, -0.000100, 0.000000, -3.141593, 0.000000],accel_mss,speed_ms,0,0.001)
  movel(p[0.453542, -0.098431, -0.000100, 0.000000, -3.141593, 0.000000],accel_mss,speed_ms,0,0.001)
  movel(p[0.450851, -0.098413, -0.000100, 0.000000, -3.141593, 0.000000],accel_mss,speed_ms,0,blend_radius_m)
  movel(p[0.448817, -0.098341, -0.000100, 0.000000, -3.141593, 0.000000],accel_mss,speed_ms,0,0.001)
  movel(p[0.447744, -0.098287, -0.000100, 0.000000, -3.141593, 0.000000],accel_mss,speed_ms,0,0.000)
  movel(p[0.446941, -0.098218, -0.000100, 0.000000, -3.141593, 0.000000],accel_mss,speed_ms,0,0.000)
  movel(p[0.446062, -0.098107, -0.000100, 0.000000, -3.141593, 0.000000],accel_mss,speed_ms,0,0.000)
  movel(p[0.445458, -0.098001, -0.000100, 0.000000, -3.141593, 0.000000],accel_mss,speed_ms,0,0.000)
  movel(p[0.444830, -0.097854, -0.000100, 0.000000, -3.141593, 0.000000],accel_mss,speed_ms,0,0.000)
  movel(p[0.444280, -0.097696, -0.000100, 0.000000, -3.141593, 0.000000],accel_mss,speed_ms,0,0.000)
  movel(p[0.444026, -0.097573, -0.000100, 0.000000, -3.141593, 0.000000],accel_mss,speed_ms,0,0.000)
  movel(p[0.443926, -0.097518, -0.000100, 0.000000, -3.141593, 0.000000],accel_mss,speed_ms,0,0.000)
  movel(p[0.443677, -0.097420, -0.000100, 0.000000, -3.141593, 0.000000],accel_mss,speed_ms,0,0.000)
  movel(p[0.443378, -0.097310, -0.000100, 0.000000, -3.141593, 0.000000],accel_mss,speed_ms,0,0.000)
  movel(p[0.443051, -0.097199, -0.000100, 0.000000, -3.141593, 0.000000],accel_mss,speed_ms,0,0.000)
  movel(p[0.442361, -0.096941, -0.000100, 0.000000, -3.141593, 0.000000],accel_mss,speed_ms,0,0.000)
  movel(p[0.441563, -0.096580, -0.000100, 0.000000, -3.141593, 0.000000],accel_mss,speed_ms,0,0.000)
  movel(p[0.440833, -0.096205, -0.000100, 0.000000, -3.141593, 0.000000],accel_mss,speed_ms,0,0.000)
  movel(p[0.440422, -0.095926, -0.000100, 0.000000, -3.141593, 0.000000],accel_mss,speed_ms,0,0.000)
  movel(p[0.440337, -0.095863, -0.000100, 0.000000, -3.141593, 0.000000],accel_mss,speed_ms,0,0.000)
  movel(p[0.440220, -0.095828, -0.000100, 0.000000, -3.141593, 0.000000],accel_mss,speed_ms,0,0.000)
  movel(p[0.440013, -0.095781, -0.000100, 0.000000, -3.141593, 0.000000],accel_mss,speed_ms,0,0.000)
  movel(p[0.439808, -0.095640, -0.000100, 0.000000, -3.141593, 0.000000],accel_mss,speed_ms,0,0.000)
  movel(p[0.439563, -0.095451, -0.000100, 0.000000, -3.141593, 0.000000],accel_mss,speed_ms,0,0.000)
  movel(p[0.439280, -0.095236, -0.000100, 0.000000, -3.141593, 0.000000],accel_mss,speed_ms,0,0.000)
  movel(p[0.438958, -0.095016, -0.000100, 0.000000, -3.141593, 0.000000],accel_mss,speed_ms,0,0.000)
  movel(p[0.438645, -0.094822, -0.000100, 0.000000, -3.141593, 0.000000],accel_mss,speed_ms,0,0.000)
  movel(p[0.438398, -0.094692, -0.000100, 0.000000, -3.141593, 0.000000],accel_mss,speed_ms,0,0.000)
  movel(p[0.438170, -0.094571, -0.000100, 0.000000, -3.141593, 0.000000],accel_mss,speed_ms,0,0.000)
  movel(p[0.437920, -0.094407, -0.000100, 0.000000, -3.141593, 0.000000],accel_mss,speed_ms,0,0.000)
  movel(p[0.437686, -0.094229, -0.000100, 0.000000, -3.141593, 0.000000],accel_mss,speed_ms,0,0.000)
  movel(p[0.437510, -0.094064, -0.000100, 0.000000, -3.141593, 0.000000],accel_mss,speed_ms,0,0.000)
  movel(p[0.437358, -0.093916, -0.000100, 0.000000, -3.141593, 0.000000],accel_mss,speed_ms,0,0.000)
  movel(p[0.437200, -0.093792, -0.000100, 0.000000, -3.141593, 0.000000],accel_mss,speed_ms,0,0.000)
  movel(p[0.437057, -0.093703, -0.000100, 0.000000, -3.141593, 0.000000],accel_mss,speed_ms,0,0.000)
  movel(p[0.436679, -0.093563, -0.000100, 0.000000, -3.141593, 0.000000],accel_mss,speed_ms,0,0.000)
  movel(p[0.434958, -0.091864, -0.000100, 0.000000, -3.141593, 0.000000],accel_mss,speed_ms,0,0.001)
  movel(p[0.433324, -0.090219, -0.000100, 0.000000, -3.141593, 0.000000],accel_mss,speed_ms,0,0.001)
  movel(p[0.432985, -0.089726, -0.000100, 0.000000, 3.141593, 0.000000],accel_mss,speed_ms,0,0.000)
  movel(p[0.432815, -0.089381, -0.000100, 0.000000, 3.141593, 0.000000],accel_mss,speed_ms,0,0.000)
  movel(p[0.432624, -0.089037, -0.000100, 0.000000, -3.141593, 0.000000],accel_mss,speed_ms,0,0.000)
  movel(p[0.432425, -0.088724, -0.000100, 0.000000, -3.141593, 0.000000],accel_mss,speed_ms,0,0.000)
  movel(p[0.432237, -0.088467, -0.000100, 0.000000, -3.141593, 0.000000],accel_mss,speed_ms,0,0.000)
  movel(p[0.431544, -0.087399, -0.000100, 0.000000, -3.141593, 0.000000],accel_mss,speed_ms,0,0.001)
  movel(p[0.430803, -0.085807, -0.000100, 0.000000, -3.141593, 0.000000],accel_mss,speed_ms,0,0.001)
  movel(p[0.430127, -0.083995, -0.000100, 0.000000, -3.141593, 0.000000],accel_mss,speed_ms,0,0.001)
  movel(p[0.429621, -0.082204, -0.000100, 0.000000, 3.141593, 0.000000],accel_mss,speed_ms,0,0.001)
  movel(p[0.429439, -0.080995, -0.000100, 0.000000, -3.141593, 0.000000],accel_mss,speed_ms,0,0.000)
  movel(p[0.429335, -0.078879, -0.000100, 0.000000, -3.141593, 0.000000],accel_mss,speed_ms,0,0.001)
  movel(p[0.429279, -0.076622, -0.000100, 0.000000, -3.141593, 0.000000],accel_mss,speed_ms,0,0.001)
  movel(p[0.429438, -0.076331, -0.000100, 0.000000, -3.141593, 0.000000],accel_mss,speed_ms,0,0.000)
  movel(p[0.429744, -0.076473, -0.000100, 0.000000, 3.141593, 0.000000],accel_mss,speed_ms,0,0.000)
  movel(p[0.430003, -0.076677, -0.000100, 0.000000, -3.141593, 0.000000],accel_mss,speed_ms,0,0.000)
  movel(p[0.430283, -0.076936, -0.000100, 0.000000, -3.141593, 0.000000],accel_mss,speed_ms,0,0.000)
  movel(p[0.430563, -0.077202, -0.000100, 0.000000, -3.141593, 0.000000],accel_mss,speed_ms,0,0.000)
  movel(p[0.430824, -0.077425, -0.000100, 0.000000, -3.141593, 0.000000],accel_mss,speed_ms,0,0.000)
  movel(p[0.431047, -0.077599, -0.000100, 0.000000, -3.141593, 0.000000],accel_mss,speed_ms,0,0.000)
  movel(p[0.431225, -0.077657, -0.000100, 0.000000, -3.141593, 0.000000],accel_mss,speed_ms,0,0.000)
  movel(p[0.431417, -0.077805, -0.000100, 0.000000, -3.141593, 0.000000],accel_mss,speed_ms,0,0.000)
  movel(p[0.431640, -0.077999, -0.000100, 0.000000, -3.141593, 0.000000],accel_mss,speed_ms,0,0.000)
  movel(p[0.431876, -0.078229, -0.000100, 0.000000, -3.141593, 0.000000],accel_mss,speed_ms,0,0.000)
  movel(p[0.432110, -0.078459, -0.000100, 0.000000, -3.141593, 0.000000],accel_mss,speed_ms,0,0.000)
  movel(p[0.432329, -0.078653, -0.000100, 0.000000, -3.141593, 0.000000],accel_mss,speed_ms,0,0.000)
  movel(p[0.432516, -0.078802, -0.000100, 0.000000, -3.141593, 0.000000],accel_mss,speed_ms,0,0.000)
  movel(p[0.432678, -0.078855, -0.000100, 0.000000, -3.141593, 0.000000],accel_mss,speed_ms,0,0.000)
  movel(p[0.432921, -0.079027, -0.000100, 0.000000, -3.141593, 0.000000],accel_mss,speed_ms,0,0.000)
  movel(p[0.433205, -0.079245, -0.000100, 0.000000, -3.141593, 0.000000],accel_mss,speed_ms,0,0.000)
  movel(p[0.433518, -0.079504, -0.000100, 0.000000, -3.141593, 0.000000],accel_mss,speed_ms,0,0.000)
  movel(p[0.433831, -0.079763, -0.000100, 0.000000, -3.141593, 0.000000],accel_mss,speed_ms,0,0.000)
  movel(p[0.434119, -0.079981, -0.000100, 0.000000, -3.141593, 0.000000],accel_mss,speed_ms,0,0.000)
  movel(p[0.434365, -0.080151, -0.000100, 0.000000, -3.141593, 0.000000],accel_mss,speed_ms,0,0.000)
  movel(p[0.434531, -0.080198, -0.000100, 0.000000, -3.141593, 0.000000],accel_mss,speed_ms,0,0.000)
  movel(p[0.434640, -0.080267, -0.000100, 0.000000, -3.141593, 0.000000],accel_mss,speed_ms,0,0.000)
  movel(p[0.434761, -0.080364, -0.000100, 0.000000, 3.141593, 0.000000],accel_mss,speed_ms,0,0.000)
  movel(p[0.434876, -0.080479, -0.000100, 0.000000, -3.141593, 0.000000],accel_mss,speed_ms,0,0.000)
  movel(p[0.434993, -0.080594, -0.000100, 0.000000, -3.141593, 0.000000],accel_mss,speed_ms,0,0.000)
  movel(p[0.435120, -0.080691, -0.000100, 0.000000, -3.141593, 0.000000],accel_mss,speed_ms,0,0.000)
  movel(p[0.435239, -0.080759, -0.000100, 0.000000, -3.141593, 0.000000],accel_mss,speed_ms,0,0.000)
  movel(p[0.435413, -0.080799, -0.000100, 0.000000, -3.141593, 0.000000],accel_mss,speed_ms,0,0.000)
  movel(p[0.435532, -0.080867, -0.000100, 0.000000, -3.141593, 0.000000],accel_mss,speed_ms,0,0.000)
  movel(p[0.435659, -0.080965, -0.000100, 0.000000, -3.141593, 0.000000],accel_mss,speed_ms,0,0.000)
  movel(p[0.435776, -0.081080, -0.000100, 0.000000, 3.141593, 0.000000],accel_mss,speed_ms,0,0.000)
  movel(p[0.435886, -0.081190, -0.000100, 0.000000, -3.141593, 0.000000],accel_mss,speed_ms,0,0.000)
  movel(p[0.435989, -0.081272, -0.000100, 0.000000, -3.141593, 0.000000],accel_mss,speed_ms,0,0.000)
  movel(p[0.436119, -0.081311, -0.000100, 0.000000, -3.141593, 0.000000],accel_mss,speed_ms,0,0.000)
  movel(p[0.436350, -0.081408, -0.000100, 0.000000, -3.141593, 0.000000],accel_mss,speed_ms,0,0.000)
  movel(p[0.436565, -0.081554, -0.000100, 0.000000, -3.141593, 0.000000],accel_mss,speed_ms,0,0.000)
  movel(p[0.436807, -0.081741, -0.000100, 0.000000, -3.141593, 0.000000],accel_mss,speed_ms,0,0.000)
  movel(p[0.437072, -0.081941, -0.000100, 0.000000, -3.141593, 0.000000],accel_mss,speed_ms,0,0.000)
  movel(p[0.437354, -0.082128, -0.000100, 0.000000, -3.141593, 0.000000],accel_mss,speed_ms,0,0.000)
  movel(p[0.437615, -0.082277, -0.000100, 0.000000, -3.141593, 0.000000],accel_mss,speed_ms,0,0.000)
  movel(p[0.437801, -0.082353, -0.000100, 0.000000, -3.141593, 0.000000],accel_mss,speed_ms,0,0.000)
  movel(p[0.437961, -0.082410, -0.000100, 0.000000, -3.141593, 0.000000],accel_mss,speed_ms,0,0.000)
  movel(p[0.438132, -0.082487, -0.000100, 0.000000, -3.141593, 0.000000],accel_mss,speed_ms,0,0.000)
  movel(p[0.438288, -0.082573, -0.000100, 0.000000, -3.141593, 0.000000],accel_mss,speed_ms,0,0.000)
  movel(p[0.438401, -0.082653, -0.000100, 0.000000, -3.141593, 0.000000],accel_mss,speed_ms,0,0.000)
  movel(p[0.438778, -0.082900, -0.000100, 0.000000, -3.141593, 0.000000],accel_mss,speed_ms,0,0.000)
  movel(p[0.440324, -0.083659, -0.000100, 0.000000, -3.141593, 0.000000],accel_mss,speed_ms,0,0.001)
  movel(p[0.441823, -0.084373, -0.000100, 0.000000, 3.141593, 0.000000],accel_mss,speed_ms,0,0.001)
  movel(p[0.442676, -0.084730, -0.000100, 0.000000, -3.141593, 0.000000],accel_mss,speed_ms,0,0.000)
  movel(p[0.442977, -0.084843, -0.000100, 0.000000, -3.141593, 0.000000],accel_mss,speed_ms,0,0.000)
  movel(p[0.443408, -0.085005, -0.000100, 0.000000, -3.141593, 0.000000],accel_mss,speed_ms,0,0.000)
  movel(p[0.443880, -0.085183, -0.000100, 0.000000, -3.141593, 0.000000],accel_mss,speed_ms,0,0.000)
  movel(p[0.444326, -0.085353, -0.000100, 0.000000, -3.141593, 0.000000],accel_mss,speed_ms,0,0.000)
  movel(p[0.444755, -0.085510, -0.000100, 0.000000, -3.141593, 0.000000],accel_mss,speed_ms,0,0.000)
  movel(p[0.445177, -0.085652, -0.000100, 0.000000, -3.141593, 0.000000],accel_mss,speed_ms,0,0.000)
  movel(p[0.445542, -0.085764, -0.000100, 0.000000, -3.141593, 0.000000],accel_mss,speed_ms,0,0.000)
  movel(p[0.445751, -0.085811, -0.000100, 0.000000, 3.141593, 0.000000],accel_mss,speed_ms,0,0.000)
  movel(p[0.445986, -0.085853, -0.000100, 0.000000, -3.141593, 0.000000],accel_mss,speed_ms,0,0.000)
  movel(p[0.446544, -0.085967, -0.000100, 0.000000, -3.141593, 0.000000],accel_mss,speed_ms,0,0.000)
  movel(p[0.447209, -0.086107, -0.000100, 0.000000, -3.141593, 0.000000],accel_mss,speed_ms,0,0.000)
  movel(p[0.447926, -0.086261, -0.000100, 0.000000, -3.141593, 0.000000],accel_mss,speed_ms,0,0.000)
  movel(p[0.449715, -0.086551, -0.000100, 0.000000, -3.141593, 0.000000],accel_mss,speed_ms,0,0.001)
  movel(p[0.451675, -0.086677, -0.000100, 0.000000, -3.141593, 0.000000],accel_mss,speed_ms,0,0.001)
  movel(p[0.453563, -0.086637, -0.000100, 0.000000, -3.141593, 0.000000],accel_mss,speed_ms,0,0.001)
  movel(p[0.455126, -0.086419, -0.000100, 0.000000, -3.141593, 0.000000],accel_mss,speed_ms,0,0.001)
  movel(p[0.457203, -0.085876, -0.000100, 0.000000, -3.141593, 0.000000],accel_mss,speed_ms,0,0.001)
  movel(p[0.459217, -0.085157, -0.000100, 0.000000, -3.141593, 0.000000],accel_mss,speed_ms,0,0.001)
  movel(p[0.460964, -0.084348, -0.000100, 0.000000, -3.141593, 0.000000],accel_mss,speed_ms,0,0.001)
  movel(p[0.462201, -0.083536, -0.000100, 0.000000, -3.141593, 0.000000],accel_mss,speed_ms,0,0.001)
  movel(p[0.462450, -0.083342, -0.000100, 0.000000, -3.141593, 0.000000],accel_mss,speed_ms,0,0.000)
  movel(p[0.462681, -0.083178, -0.000100, 0.000000, -3.141593, 0.000000],accel_mss,speed_ms,0,0.000)
  movel(p[0.462878, -0.083051, -0.000100, 0.000000, -3.141593, 0.000000],accel_mss,speed_ms,0,0.000)
  movel(p[0.463036, -0.083002, -0.000100, 0.000000, -3.141593, 0.000000],accel_mss,speed_ms,0,0.000)
  movel(p[0.463244, -0.082831, -0.000100, 0.000000, -3.141593, 0.000000],accel_mss,speed_ms,0,0.000)
  movel(p[0.463487, -0.082613, -0.000100, 0.000000, -3.141593, 0.000000],accel_mss,speed_ms,0,0.000)
  movel(p[0.463751, -0.082354, -0.000100, 0.000000, -3.141593, 0.000000],accel_mss,speed_ms,0,0.000)
  movel(p[0.464016, -0.082095, -0.000100, 0.000000, -3.141593, 0.000000],accel_mss,speed_ms,0,0.000)
  movel(p[0.464263, -0.081877, -0.000100, 0.000000, -3.141593, 0.000000],accel_mss,speed_ms,0,0.000)
  movel(p[0.464476, -0.081709, -0.000100, 0.000000, -3.141593, 0.000000],accel_mss,speed_ms,0,0.000)
  movel(p[0.464803, -0.081582, -0.000100, 0.000000, -3.141593, 0.000000],accel_mss,speed_ms,0,0.000)
  movel(p[0.465885, -0.080516, -0.000100, 0.000000, -3.141593, 0.000000],accel_mss,speed_ms,0,0.001)
  movel(p[0.466954, -0.079438, -0.000100, 0.000000, -3.141593, 0.000000],accel_mss,speed_ms,0,0.001)
  movel(p[0.467051, -0.079201, -0.000100, 0.000000, -3.141593, 0.000000],accel_mss,speed_ms,0,0.000)
  movel(p[0.467249, -0.078894, -0.000100, 0.000000, -3.141593, 0.000000],accel_mss,speed_ms,0,0.000)
  movel(p[0.467467, -0.078644, -0.000100, 0.000000, -3.141593, 0.000000],accel_mss,speed_ms,0,0.000)
  movel(p[0.467726, -0.078379, -0.000100, 0.000000, -3.141593, 0.000000],accel_mss,speed_ms,0,0.000)
  movel(p[0.467984, -0.078116, -0.000100, 0.000000, -3.141593, 0.000000],accel_mss,speed_ms,0,0.000)
  movel(p[0.468202, -0.077873, -0.000100, 0.000000, -3.141593, 0.000000],accel_mss,speed_ms,0,0.000)
  movel(p[0.468373, -0.077665, -0.000100, 0.000000, -3.141593, 0.000000],accel_mss,speed_ms,0,0.000)
  movel(p[0.468424, -0.077507, -0.000100, 0.000000, -3.141593, 0.000000],accel_mss,speed_ms,0,0.000)
  movel(p[0.468571, -0.077290, -0.000100, 0.000000, -3.141593, 0.000000],accel_mss,speed_ms,0,0.000)
  movel(p[0.468759, -0.077034, -0.000100, 0.000000, -3.141593, 0.000000],accel_mss,speed_ms,0,0.000)
  movel(p[0.468981, -0.076756, -0.000100, 0.000000, -3.141593, 0.000000],accel_mss,speed_ms,0,0.000)
  movel(p[0.469643, -0.075853, -0.000100, 0.000000, -3.141593, 0.000000],accel_mss,speed_ms,0,0.000)
  movel(p[0.470391, -0.074620, -0.000100, 0.000000, -3.141593, 0.000000],accel_mss,speed_ms,0,0.001)
  movel(p[0.471130, -0.073237, -0.000100, 0.000000, -3.141593, 0.000000],accel_mss,speed_ms,0,0.001)
  movel(p[0.471773, -0.071854, -0.000100, 0.000000, -3.141593, 0.000000],accel_mss,speed_ms,0,0.001)
  movel(p[0.471892, -0.071581, -0.000100, 0.000000, -3.141593, 0.000000],accel_mss,speed_ms,0,0.000)
  movel(p[0.472037, -0.071254, -0.000100, 0.000000, -3.141593, 0.000000],accel_mss,speed_ms,0,0.000)
  movel(p[0.472185, -0.070927, -0.000100, 0.000000, -3.141593, 0.000000],accel_mss,speed_ms,0,0.000)
  movel(p[0.472311, -0.070654, -0.000100, 0.000000, -3.141593, 0.000000],accel_mss,speed_ms,0,0.000)
  movel(p[0.472422, -0.070402, -0.000100, 0.000000, -3.141593, 0.000000],accel_mss,speed_ms,0,0.000)
  movel(p[0.472525, -0.070142, -0.000100, 0.000000, -3.141593, 0.000000],accel_mss,speed_ms,0,0.000)
  movel(p[0.472606, -0.069909, -0.000100, 0.000000, -3.141593, 0.000000],accel_mss,speed_ms,0,0.000)
  movel(p[0.472645, -0.069754, -0.000100, 0.000000, 3.141593, 0.000000],accel_mss,speed_ms,0,0.000)
  movel(p[0.472687, -0.069571, -0.000100, 0.000000, -3.141593, 0.000000],accel_mss,speed_ms,0,0.000)
  movel(p[0.472798, -0.069168, -0.000100, 0.000000, -3.141593, 0.000000],accel_mss,speed_ms,0,0.000)
  movel(p[0.472935, -0.068689, -0.000100, 0.000000, -3.141593, 0.000000],accel_mss,speed_ms,0,0.000)
  movel(p[0.473087, -0.068179, -0.000100, 0.000000, -3.141593, 0.000000],accel_mss,speed_ms,0,0.000)
  movel(p[0.473524, -0.066608, -0.000100, 0.000000, -3.141593, 0.000000],accel_mss,speed_ms,0,0.001)
  movel(p[0.473759, -0.065410, -0.000100, 0.000000, -3.141593, 0.000000],accel_mss,speed_ms,0,0.000)
  movel(p[0.473902, -0.063985, -0.000100, 0.000000, -3.141593, 0.000000],accel_mss,speed_ms,0,0.001)
  movel(p[0.474040, -0.061391, -0.000100, 0.000000, -3.141593, 0.000000],accel_mss,speed_ms,0,blend_radius_m)
  movel(p[0.474099, -0.059732, -0.000100, 0.000000, -3.141593, 0.000000],accel_mss,speed_ms,0,0.001)
  movel(p[0.474028, -0.059142, -0.000100, 0.000000, -3.141593, 0.000000],accel_mss,speed_ms,0,0.000)
  movel(p[0.473853, -0.059106, -0.000100, 0.000000, -3.141593, 0.000000],accel_mss,speed_ms,0,0.000)
  movel(p[0.473555, -0.059591, -0.000100, 0.000000, -3.141593, 0.000000],accel_mss,speed_ms,0,0.000)
  movel(p[0.473427, -0.059845, -0.000100, 0.000000, 3.141593, 0.000000],accel_mss,speed_ms,0,0.000)
  movel(p[0.473254, -0.060143, -0.000100, 0.000000, -3.141593, 0.000000],accel_mss,speed_ms,0,0.000)
  movel(p[0.473066, -0.060437, -0.000100, 0.000000, -3.141593, 0.000000],accel_mss,speed_ms,0,0.000)
  movel(p[0.472893, -0.060679, -0.000100, 0.000000, -3.141593, 0.000000],accel_mss,speed_ms,0,0.000)
  movel(p[0.472731, -0.060907, -0.000100, 0.000000, 3.141593, 0.000000],accel_mss,speed_ms,0,0.000)
  movel(p[0.472576, -0.061160, -0.000100, 0.000000, 3.141593, 0.000000],accel_mss,speed_ms,0,0.000)
  movel(p[0.472448, -0.061399, -0.000100, 0.000000, -3.141593, 0.000000],accel_mss,speed_ms,0,0.000)
  movel(p[0.472377, -0.061579, -0.000100, 0.000000, -3.141593, 0.000000],accel_mss,speed_ms,0,0.000)
  movel(p[0.472322, -0.061737, -0.000100, 0.000000, -3.141593, 0.000000],accel_mss,speed_ms,0,0.000)
  movel(p[0.472249, -0.061904, -0.000100, 0.000000, -3.141593, 0.000000],accel_mss,speed_ms,0,0.000)
  movel(p[0.472171, -0.062053, -0.000100, 0.000000, -3.141593, 0.000000],accel_mss,speed_ms,0,0.000)
  movel(p[0.472101, -0.062157, -0.000100, 0.000000, -3.141593, 0.000000],accel_mss,speed_ms,0,0.000)
  movel(p[0.471944, -0.062372, -0.000100, 0.000000, -3.141593, 0.000000],accel_mss,speed_ms,0,0.000)
  movel(p[0.471762, -0.062663, -0.000100, 0.000000, -3.141593, 0.000000],accel_mss,speed_ms,0,0.000)
  movel(p[0.471555, -0.063022, -0.000100, 0.000000, -3.141593, 0.000000],accel_mss,speed_ms,0,0.000)
  movel(p[0.471325, -0.063454, -0.000100, 0.000000, -3.141593, 0.000000],accel_mss,speed_ms,0,0.000)
  movel(p[0.471214, -0.063659, -0.000100, 0.000000, -3.141593, 0.000000],accel_mss,speed_ms,0,0.000)
  movel(p[0.471074, -0.063904, -0.000100, 0.000000, -3.141593, 0.000000],accel_mss,speed_ms,0,0.000)
  movel(p[0.470929, -0.064149, -0.000100, 0.000000, -3.141593, 0.000000],accel_mss,speed_ms,0,0.000)
  movel(p[0.470801, -0.064354, -0.000100, 0.000000, -3.141593, 0.000000],accel_mss,speed_ms,0,0.000)
  movel(p[0.470673, -0.064559, -0.000100, 0.000000, 3.141593, 0.000000],accel_mss,speed_ms,0,0.000)
  movel(p[0.470528, -0.064804, -0.000100, 0.000000, -3.141593, 0.000000],accel_mss,speed_ms,0,0.000)
  movel(p[0.470389, -0.065049, -0.000100, 0.000000, -3.141593, 0.000000],accel_mss,speed_ms,0,0.000)
  movel(p[0.470281, -0.065254, -0.000100, 0.000000, -3.141593, 0.000000],accel_mss,speed_ms,0,0.000)
  movel(p[0.470172, -0.065459, -0.000100, 0.000000, 3.141593, 0.000000],accel_mss,speed_ms,0,0.000)
  movel(p[0.470032, -0.065704, -0.000100, 0.000000, -3.141593, 0.000000],accel_mss,speed_ms,0,0.000)
  movel(p[0.469887, -0.065949, -0.000100, 0.000000, -3.141593, 0.000000],accel_mss,speed_ms,0,0.000)
  movel(p[0.469758, -0.066154, -0.000100, 0.000000, -3.141593, 0.000000],accel_mss,speed_ms,0,0.000)
  movel(p[0.469626, -0.066364, -0.000100, 0.000000, -3.141593, 0.000000],accel_mss,speed_ms,0,0.000)
  movel(p[0.469473, -0.066626, -0.000100, 0.000000, -3.141593, 0.000000],accel_mss,speed_ms,0,0.000)
  movel(p[0.469323, -0.066895, -0.000100, 0.000000, -3.141593, 0.000000],accel_mss,speed_ms,0,0.000)
  movel(p[0.469202, -0.067129, -0.000100, 0.000000, -3.141593, 0.000000],accel_mss,speed_ms,0,0.000)
  movel(p[0.468991, -0.067527, -0.000100, 0.000000, -3.141593, 0.000000],accel_mss,speed_ms,0,0.000)
  movel(p[0.468690, -0.068054, -0.000100, 0.000000, -3.141593, 0.000000],accel_mss,speed_ms,0,0.000)
  movel(p[0.468309, -0.068696, -0.000100, 0.000000, -3.141593, 0.000000],accel_mss,speed_ms,0,0.000)
  movel(p[0.467842, -0.069458, -0.000100, 0.000000, -3.141593, 0.000000],accel_mss,speed_ms,0,0.000)
  movel(p[0.467754, -0.069607, -0.000100, 0.000000, -3.141593, 0.000000],accel_mss,speed_ms,0,0.000)
  movel(p[0.467637, -0.069821, -0.000100, 0.000000, -3.141593, 0.000000],accel_mss,speed_ms,0,0.000)
  movel(p[0.467513, -0.070056, -0.000100, 0.000000, -3.141593, 0.000000],accel_mss,speed_ms,0,0.000)
  movel(p[0.467401, -0.070279, -0.000100, 0.000000, -3.141593, 0.000000],accel_mss,speed_ms,0,0.000)
  movel(p[0.467279, -0.070513, -0.000100, 0.000000, -3.141593, 0.000000],accel_mss,speed_ms,0,0.000)
  movel(p[0.467124, -0.070782, -0.000100, 0.000000, -3.141593, 0.000000],accel_mss,speed_ms,0,0.000)
  movel(p[0.466962, -0.071044, -0.000100, 0.000000, -3.141593, 0.000000],accel_mss,speed_ms,0,0.000)
  movel(p[0.466819, -0.071254, -0.000100, 0.000000, -3.141593, 0.000000],accel_mss,speed_ms,0,0.000)
  movel(p[0.466688, -0.071443, -0.000100, 0.000000, -3.141593, 0.000000],accel_mss,speed_ms,0,0.000)
  movel(p[0.466561, -0.071638, -0.000100, 0.000000, -3.141593, 0.000000],accel_mss,speed_ms,0,0.000)
  movel(p[0.466455, -0.071813, -0.000100, 0.000000, -3.141593, 0.000000],accel_mss,speed_ms,0,0.000)
  movel(p[0.466396, -0.071929, -0.000100, 0.000000, -3.141593, 0.000000],accel_mss,speed_ms,0,0.000)
  movel(p[0.466339, -0.072045, -0.000100, 0.000000, -3.141593, 0.000000],accel_mss,speed_ms,0,0.000)
  movel(p[0.466240, -0.072220, -0.000100, 0.000000, -3.141593, 0.000000],accel_mss,speed_ms,0,0.000)
  movel(p[0.466123, -0.072415, -0.000100, 0.000000, -3.141593, 0.000000],accel_mss,speed_ms,0,0.000)
  movel(p[0.466004, -0.072604, -0.000100, 0.000000, -3.141593, 0.000000],accel_mss,speed_ms,0,0.000)
  movel(p[0.465876, -0.072809, -0.000100, 0.000000, -3.141593, 0.000000],accel_mss,speed_ms,0,0.000)
  movel(p[0.465736, -0.073054, -0.000100, 0.000000, -3.141593, 0.000000],accel_mss,speed_ms,0,0.000)
  movel(p[0.465604, -0.073299, -0.000100, 0.000000, 3.141593, 0.000000],accel_mss,speed_ms,0,0.000)
  movel(p[0.465504, -0.073504, -0.000100, 0.000000, -3.141593, 0.000000],accel_mss,speed_ms,0,0.000)
  movel(p[0.465406, -0.073692, -0.000100, 0.000000, -3.141593, 0.000000],accel_mss,speed_ms,0,0.000)
  movel(p[0.465283, -0.073884, -0.000100, 0.000000, -3.141593, 0.000000],accel_mss,speed_ms,0,0.000)
  movel(p[0.465154, -0.074053, -0.000100, 0.000000, -3.141593, 0.000000],accel_mss,speed_ms,0,0.000)
  movel(p[0.465041, -0.074166, -0.000100, 0.000000, -3.141593, 0.000000],accel_mss,speed_ms,0,0.000)
  movel(p[0.464924, -0.074289, -0.000100, 0.000000, -3.141593, 0.000000],accel_mss,speed_ms,0,0.000)
  movel(p[0.464778, -0.074497, -0.000100, 0.000000, -3.141593, 0.000000],accel_mss,speed_ms,0,0.000)
  movel(p[0.464631, -0.074743, -0.000100, 0.000000, -3.141593, 0.000000],accel_mss,speed_ms,0,0.000)
  movel(p[0.464505, -0.074995, -0.000100, 0.000000, -3.141593, 0.000000],accel_mss,speed_ms,0,0.000)
  movel(p[0.464374, -0.075251, -0.000100, 0.000000, -3.141593, 0.000000],accel_mss,speed_ms,0,0.000)
  movel(p[0.464215, -0.075513, -0.000100, 0.000000, -3.141593, 0.000000],accel_mss,speed_ms,0,0.000)
  movel(p[0.464051, -0.075742, -0.000100, 0.000000, -3.141593, 0.000000],accel_mss,speed_ms,0,0.000)
  movel(p[0.463912, -0.075893, -0.000100, 0.000000, -3.141593, 0.000000],accel_mss,speed_ms,0,0.000)
  movel(p[0.463793, -0.076012, -0.000100, 0.000000, -3.141593, 0.000000],accel_mss,speed_ms,0,0.000)
  movel(p[0.463692, -0.076136, -0.000100, 0.000000, -3.141593, 0.000000],accel_mss,speed_ms,0,0.000)
  movel(p[0.463620, -0.076248, -0.000100, 0.000000, -3.141593, 0.000000],accel_mss,speed_ms,0,0.000)
  movel(p[0.463571, -0.076416, -0.000100, 0.000000, -3.141593, 0.000000],accel_mss,speed_ms,0,0.000)
  movel(p[0.463358, -0.076703, -0.000100, 0.000000, -3.141593, 0.000000],accel_mss,speed_ms,0,0.000)
  movel(p[0.463092, -0.077040, -0.000100, 0.000000, -3.141593, 0.000000],accel_mss,speed_ms,0,0.000)
  movel(p[0.462776, -0.077410, -0.000100, 0.000000, -3.141593, 0.000000],accel_mss,speed_ms,0,0.000)
  movel(p[0.462460, -0.077780, -0.000100, 0.000000, -3.141593, 0.000000],accel_mss,speed_ms,0,0.000)
  movel(p[0.462193, -0.078114, -0.000100, 0.000000, -3.141593, 0.000000],accel_mss,speed_ms,0,0.000)
  movel(p[0.461979, -0.078400, -0.000100, 0.000000, -3.141593, 0.000000],accel_mss,speed_ms,0,0.000)
  movel(p[0.461877, -0.078662, -0.000100, 0.000000, -3.141593, 0.000000],accel_mss,speed_ms,0,0.000)
  movel(p[0.461414, -0.079096, -0.000100, 0.000000, -3.141593, 0.000000],accel_mss,speed_ms,0,0.000)
  movel(p[0.460935, -0.079508, -0.000100, 0.000000, -3.141593, 0.000000],accel_mss,speed_ms,0,0.000)
  movel(p[0.460736, -0.079579, -0.000100, 0.000000, -3.141593, 0.000000],accel_mss,speed_ms,0,0.000)
  movel(p[0.460640, -0.079634, -0.000100, 0.000000, -3.141593, 0.000000],accel_mss,speed_ms,0,0.000)
  movel(p[0.460599, -0.079766, -0.000100, 0.000000, -3.141593, 0.000000],accel_mss,speed_ms,0,0.000)
  movel(p[0.460500, -0.079947, -0.000100, 0.000000, -3.141593, 0.000000],accel_mss,speed_ms,0,0.000)
  movel(p[0.460391, -0.080042, -0.000100, 0.000000, -3.141593, 0.000000],accel_mss,speed_ms,0,0.000)
  movel(p[0.460262, -0.080119, -0.000100, 0.000000, -3.141593, 0.000000],accel_mss,speed_ms,0,0.000)
  movel(p[0.460092, -0.080204, -0.000100, 0.000000, -3.141593, 0.000000],accel_mss,speed_ms,0,0.000)
  movel(p[0.459848, -0.080328, -0.000100, 0.000000, -3.141593, 0.000000],accel_mss,speed_ms,0,0.000)
  movel(p[0.459580, -0.080466, -0.000100, 0.000000, -3.141593, 0.000000],accel_mss,speed_ms,0,0.000)
  movel(p[0.459326, -0.080598, -0.000100, 0.000000, -3.141593, 0.000000],accel_mss,speed_ms,0,0.000)
  movel(p[0.457809, -0.081341, -0.000100, 0.000000, -3.141593, 0.000000],accel_mss,speed_ms,0,0.001)
  movel(p[0.456519, -0.081859, -0.000100, 0.000000, -3.141593, 0.000000],accel_mss,speed_ms,0,0.001)
  movel(p[0.455409, -0.082175, -0.000100, 0.000000, -3.141593, 0.000000],accel_mss,speed_ms,0,0.000)
  movel(p[0.454451, -0.082292, -0.000100, 0.000000, -3.141593, 0.000000],accel_mss,speed_ms,0,0.000)
  movel(p[0.454199, -0.082302, -0.000100, 0.000000, -3.141593, 0.000000],accel_mss,speed_ms,0,0.000)
  movel(p[0.453872, -0.082323, -0.000100, 0.000000, -3.141593, 0.000000],accel_mss,speed_ms,0,0.000)
  movel(p[0.453527, -0.082351, -0.000100, 0.000000, -3.141593, 0.000000],accel_mss,speed_ms,0,0.000)
  movel(p[0.453218, -0.082380, -0.000100, 0.000000, -3.141593, 0.000000],accel_mss,speed_ms,0,0.000)
  movel(p[0.452864, -0.082418, -0.000100, 0.000000, -3.141593, 0.000000],accel_mss,speed_ms,0,0.000)
  movel(p[0.452511, -0.082456, -0.000100, 0.000000, -3.141593, 0.000000],accel_mss,speed_ms,0,0.000)
  movel(p[0.452527, -0.083115, -0.000100, 0.000000, -3.141593, 0.000000],accel_mss,speed_ms,0,0.000)
  movel(p[0.452543, -0.083775, -0.000100, 0.000000, -3.141593, 0.000000],accel_mss,speed_ms,0,0.000)
  movel(p[0.452550, -0.084486, -0.000100, 0.000000, -3.141593, 0.000000],accel_mss,speed_ms,0,0.000)
  movel(p[0.452518, -0.084900, -0.000100, 0.000000, -3.141593, 0.000000],accel_mss,speed_ms,0,0.000)
  movel(p[0.452442, -0.085177, -0.000100, 0.000000, -3.141593, 0.000000],accel_mss,speed_ms,0,0.000)
  movel(p[0.452306, -0.085394, -0.000100, 0.000000, 3.141593, 0.000000],accel_mss,speed_ms,0,0.000)
  movel(p[0.451657, -0.085809, -0.000100, 0.000000, -3.141593, 0.000000],accel_mss,speed_ms,0,0.000)
  movel(p[0.450649, -0.085992, -0.000100, 0.000000, -3.141593, 0.000000],accel_mss,speed_ms,0,0.000)
  movel(p[0.449641, -0.085930, -0.000100, 0.000000, -3.141593, 0.000000],accel_mss,speed_ms,0,0.000)
  movel(p[0.448996, -0.085591, -0.000100, 0.000000, -3.141593, 0.000000],accel_mss,speed_ms,0,0.000)
  movel(p[0.448837, -0.085388, -0.000100, 0.000000, -3.141593, 0.000000],accel_mss,speed_ms,0,0.000)
  movel(p[0.448743, -0.085167, -0.000100, 0.000000, 3.141593, 0.000000],accel_mss,speed_ms,0,0.000)
  movel(p[0.448700, -0.084875, -0.000100, 0.000000, -3.141593, 0.000000],accel_mss,speed_ms,0,0.000)
  movel(p[0.448696, -0.084432, -0.000100, 0.000000, -3.141593, 0.000000],accel_mss,speed_ms,0,0.000)
  movel(p[0.448725, -0.083960, -0.000100, 0.000000, -3.141593, 0.000000],accel_mss,speed_ms,0,0.000)
  movel(p[0.448794, -0.083661, -0.000100, 0.000000, -3.141593, 0.000000],accel_mss,speed_ms,0,0.000)
  movel(p[0.448930, -0.083414, -0.000100, 0.000000, -3.141593, 0.000000],accel_mss,speed_ms,0,0.000)
  movel(p[0.449178, -0.083132, -0.000100, 0.000000, 3.141593, 0.000000],accel_mss,speed_ms,0,0.000)
  movel(p[0.449410, -0.082901, -0.000100, 0.000000, -3.141593, 0.000000],accel_mss,speed_ms,0,0.000)
  movel(p[0.449641, -0.082669, -0.000100, 0.000000, -3.141593, 0.000000],accel_mss,speed_ms,0,0.000)
  movel(p[0.449634, -0.083021, -0.000100, 0.000000, -3.141593, 0.000000],accel_mss,speed_ms,0,0.000)
  movel(p[0.449627, -0.083373, -0.000100, 0.000000, -3.141593, 0.000000],accel_mss,speed_ms,0,0.000)
  movel(p[0.449657, -0.083877, -0.000100, 0.000000, -3.141593, 0.000000],accel_mss,speed_ms,0,0.000)
  movel(p[0.449776, -0.084236, -0.000100, 0.000000, -3.141593, 0.000000],accel_mss,speed_ms,0,0.000)
  movel(p[0.449980, -0.084450, -0.000100, 0.000000, 3.141593, 0.000000],accel_mss,speed_ms,0,0.000)
  movel(p[0.450260, -0.084529, -0.000100, 0.000000, -3.141593, 0.000000],accel_mss,speed_ms,0,0.000)
  movel(p[0.450541, -0.084430, -0.000100, 0.000000, -3.141593, 0.000000],accel_mss,speed_ms,0,0.000)
  movel(p[0.450782, -0.084151, -0.000100, 0.000000, -3.141593, 0.000000],accel_mss,speed_ms,0,0.000)
  movel(p[0.450945, -0.083736, -0.000100, 0.000000, 3.141593, 0.000000],accel_mss,speed_ms,0,0.000)
  movel(p[0.451001, -0.083251, -0.000100, 0.000000, -3.141593, 0.000000],accel_mss,speed_ms,0,0.000)
  movel(p[0.450961, -0.082796, -0.000100, 0.000000, -3.141593, 0.000000],accel_mss,speed_ms,0,0.000)
  movel(p[0.450833, -0.082501, -0.000100, 0.000000, -3.141593, 0.000000],accel_mss,speed_ms,0,0.000)
  movel(p[0.450606, -0.082336, -0.000100, 0.000000, -3.141593, 0.000000],accel_mss,speed_ms,0,0.000)
  movel(p[0.450268, -0.082279, -0.000100, 0.000000, -3.141593, 0.000000],accel_mss,speed_ms,0,0.000)
  movel(p[0.449800, -0.082207, -0.000100, 0.000000, -3.141593, 0.000000],accel_mss,speed_ms,0,0.000)
  movel(p[0.448160, -0.081683, -0.000100, 0.000000, -3.141593, 0.000000],accel_mss,speed_ms,0,0.001)
  movel(p[0.446517, -0.081136, -0.000100, 0.000000, -3.141593, 0.000000],accel_mss,speed_ms,0,0.001)
  movel(p[0.446126, -0.080926, -0.000100, 0.000000, -3.141593, 0.000000],accel_mss,speed_ms,0,0.000)
  movel(p[0.445924, -0.080791, -0.000100, 0.000000, -3.141593, 0.000000],accel_mss,speed_ms,0,0.000)
  movel(p[0.445422, -0.080502, -0.000100, 0.000000, -3.141593, 0.000000],accel_mss,speed_ms,0,0.000)
  movel(p[0.444838, -0.080177, -0.000100, 0.000000, -3.141593, 0.000000],accel_mss,speed_ms,0,0.000)
  movel(p[0.444240, -0.079858, -0.000100, 0.000000, -3.141593, 0.000000],accel_mss,speed_ms,0,0.000)
  movel(p[0.444004, -0.079718, -0.000100, 0.000000, -3.141593, 0.000000],accel_mss,speed_ms,0,0.000)
  movel(p[0.443736, -0.079527, -0.000100, 0.000000, 3.141593, 0.000000],accel_mss,speed_ms,0,0.000)
  movel(p[0.443478, -0.079320, -0.000100, 0.000000, -3.141593, 0.000000],accel_mss,speed_ms,0,0.000)
  movel(p[0.443275, -0.079128, -0.000100, 0.000000, 3.141593, 0.000000],accel_mss,speed_ms,0,0.000)
  movel(p[0.443096, -0.078956, -0.000100, 0.000000, -3.141593, 0.000000],accel_mss,speed_ms,0,0.000)
  movel(p[0.442913, -0.078811, -0.000100, 0.000000, -3.141593, 0.000000],accel_mss,speed_ms,0,0.000)
  movel(p[0.442750, -0.078706, -0.000100, 0.000000, -3.141593, 0.000000],accel_mss,speed_ms,0,0.000)
  movel(p[0.442648, -0.078679, -0.000100, 0.000000, -3.141593, 0.000000],accel_mss,speed_ms,0,0.000)
  movel(p[0.442508, -0.078611, -0.000100, 0.000000, -3.141593, 0.000000],accel_mss,speed_ms,0,0.000)
  movel(p[0.442451, -0.078449, -0.000100, 0.000000, -3.141593, 0.000000],accel_mss,speed_ms,0,0.000)
  movel(p[0.442374, -0.078259, -0.000100, 0.000000, -3.141593, 0.000000],accel_mss,speed_ms,0,0.000)
  movel(p[0.442288, -0.078178, -0.000100, 0.000000, -3.141593, 0.000000],accel_mss,speed_ms,0,0.000)
  movel(p[0.442188, -0.078125, -0.000100, 0.000000, -3.141593, 0.000000],accel_mss,speed_ms,0,0.000)
  movel(p[0.441897, -0.077965, -0.000100, 0.000000, -3.141593, 0.000000],accel_mss,speed_ms,0,0.000)
  movel(p[0.441521, -0.077641, -0.000100, 0.000000, -3.141593, 0.000000],accel_mss,speed_ms,0,0.000)
  movel(p[0.441183, -0.077292, -0.000100, 0.000000, -3.141593, 0.000000],accel_mss,speed_ms,0,0.000)
  movel(p[0.441105, -0.077093, -0.000100, 0.000000, -3.141593, 0.000000],accel_mss,speed_ms,0,0.000)
  movel(p[0.440987, -0.076872, -0.000100, 0.000000, -3.141593, 0.000000],accel_mss,speed_ms,0,0.000)
  movel(p[0.440860, -0.076719, -0.000100, 0.000000, -3.141593, 0.000000],accel_mss,speed_ms,0,0.000)
  movel(p[0.440710, -0.076568, -0.000100, 0.000000, -3.141593, 0.000000],accel_mss,speed_ms,0,0.000)
  movel(p[0.440550, -0.076406, -0.000100, 0.000000, 3.141593, 0.000000],accel_mss,speed_ms,0,0.000)
  movel(p[0.440394, -0.076223, -0.000100, 0.000000, 3.141593, 0.000000],accel_mss,speed_ms,0,0.000)
  movel(p[0.440262, -0.076044, -0.000100, 0.000000, -3.141593, 0.000000],accel_mss,speed_ms,0,0.000)
  movel(p[0.440182, -0.075904, -0.000100, 0.000000, -3.141593, 0.000000],accel_mss,speed_ms,0,0.000)
  movel(p[0.440099, -0.075731, -0.000100, 0.000000, -3.141593, 0.000000],accel_mss,speed_ms,0,0.000)
  movel(p[0.439933, -0.075406, -0.000100, 0.000000, 3.141593, 0.000000],accel_mss,speed_ms,0,0.000)
  movel(p[0.439734, -0.075024, -0.000100, 0.000000, -3.141593, 0.000000],accel_mss,speed_ms,0,0.000)
  movel(p[0.439524, -0.074629, -0.000100, 0.000000, -3.141593, 0.000000],accel_mss,speed_ms,0,0.000)
  movel(p[0.439146, -0.073851, -0.000100, 0.000000, -3.141593, 0.000000],accel_mss,speed_ms,0,0.000)
  movel(p[0.438777, -0.072947, -0.000100, 0.000000, -3.141593, 0.000000],accel_mss,speed_ms,0,0.000)
  movel(p[0.438478, -0.072083, -0.000100, 0.000000, -3.141593, 0.000000],accel_mss,speed_ms,0,0.000)
  movel(p[0.438330, -0.071457, -0.000100, 0.000000, -3.141593, 0.000000],accel_mss,speed_ms,0,0.000)
  movel(p[0.438134, -0.070061, -0.000100, 0.000000, -3.141593, 0.000000],accel_mss,speed_ms,0,0.001)
  movel(p[0.438038, -0.068930, -0.000100, 0.000000, -3.141593, 0.000000],accel_mss,speed_ms,0,0.000)
  movel(p[0.438028, -0.067856, -0.000100, 0.000000, -3.141593, 0.000000],accel_mss,speed_ms,0,0.000)
  movel(p[0.438095, -0.066649, -0.000100, 0.000000, 3.141593, 0.000000],accel_mss,speed_ms,0,0.000)
  movel(p[0.438160, -0.065909, -0.000100, 0.000000, -3.141593, 0.000000],accel_mss,speed_ms,0,0.000)
  movel(p[0.438226, -0.065214, -0.000100, 0.000000, -3.141593, 0.000000],accel_mss,speed_ms,0,0.000)
  movel(p[0.438287, -0.064628, -0.000100, 0.000000, 3.141593, 0.000000],accel_mss,speed_ms,0,0.000)
  movel(p[0.438325, -0.064354, -0.000100, 0.000000, -3.141593, 0.000000],accel_mss,speed_ms,0,0.000)
  movel(p[0.438360, -0.064144, -0.000100, 0.000000, -3.141593, 0.000000],accel_mss,speed_ms,0,0.000)
  movel(p[0.438404, -0.063882, -0.000100, 0.000000, -3.141593, 0.000000],accel_mss,speed_ms,0,0.000)
  movel(p[0.438448, -0.063613, -0.000100, 0.000000, 3.141593, 0.000000],accel_mss,speed_ms,0,0.000)
  movel(p[0.438486, -0.063379, -0.000100, 0.000000, -3.141593, 0.000000],accel_mss,speed_ms,0,0.000)
  movel(p[0.438595, -0.062866, -0.000100, 0.000000, -3.141593, 0.000000],accel_mss,speed_ms,0,0.000)
  movel(p[0.438790, -0.062183, -0.000100, 0.000000, -3.141593, 0.000000],accel_mss,speed_ms,0,0.000)
  movel(p[0.439021, -0.061477, -0.000100, 0.000000, -3.141593, 0.000000],accel_mss,speed_ms,0,0.000)
  movel(p[0.439251, -0.060881, -0.000100, 0.000000, -3.141593, 0.000000],accel_mss,speed_ms,0,0.000)
  movel(p[0.439328, -0.060694, -0.000100, 0.000000, -3.141593, 0.000000],accel_mss,speed_ms,0,0.000)
  movel(p[0.439392, -0.060522, -0.000100, 0.000000, -3.141593, 0.000000],accel_mss,speed_ms,0,0.000)
  movel(p[0.439442, -0.060378, -0.000100, 0.000000, -3.141593, 0.000000],accel_mss,speed_ms,0,0.000)
  movel(p[0.439507, -0.060074, -0.000100, 0.000000, 3.141593, 0.000000],accel_mss,speed_ms,0,0.000)
  movel(p[0.439854, -0.059365, -0.000100, 0.000000, -3.141593, 0.000000],accel_mss,speed_ms,0,0.000)
  movel(p[0.440217, -0.058672, -0.000100, 0.000000, -3.141593, 0.000000],accel_mss,speed_ms,0,0.000)
  movel(p[0.440398, -0.058452, -0.000100, 0.000000, 3.141593, 0.000000],accel_mss,speed_ms,0,0.000)
  movel(p[0.440714, -0.058287, -0.000100, 0.000000, -3.141593, 0.000000],accel_mss,speed_ms,0,0.000)
  movel(p[0.441343, -0.058143, -0.000100, 0.000000, -3.141593, 0.000000],accel_mss,speed_ms,0,0.000)
  movel(p[0.441981, -0.058044, -0.000100, 0.000000, -3.141593, 0.000000],accel_mss,speed_ms,0,0.000)
  movel(p[0.442195, -0.058117, -0.000100, 0.000000, -3.141593, 0.000000],accel_mss,speed_ms,0,0.000)
  movel(p[0.442217, -0.058215, -0.000100, 0.000000, -3.141593, 0.000000],accel_mss,speed_ms,0,0.000)
  movel(p[0.442024, -0.058701, -0.000100, 0.000000, 3.141593, 0.000000],accel_mss,speed_ms,0,0.000)
  movel(p[0.441770, -0.059279, -0.000100, 0.000000, -3.141593, 0.000000],accel_mss,speed_ms,0,0.000)
  movel(p[0.441445, -0.059944, -0.000100, 0.000000, -3.141593, 0.000000],accel_mss,speed_ms,0,0.000)
  movel(p[0.441010, -0.060799, -0.000100, 0.000000, -3.141593, 0.000000],accel_mss,speed_ms,0,0.000)
  movel(p[0.440576, -0.061654, -0.000100, 0.000000, -3.141593, 0.000000],accel_mss,speed_ms,0,0.000)
  movel(p[0.440561, -0.062929, -0.000100, 0.000000, 3.141593, 0.000000],accel_mss,speed_ms,0,0.001)
  movel(p[0.440547, -0.064204, -0.000100, 0.000000, -3.141593, 0.000000],accel_mss,speed_ms,0,0.001)
  movel(p[0.440547, -0.065235, -0.000100, 0.000000, -3.141593, 0.000000],accel_mss,speed_ms,0,0.000)
  movel(p[0.440571, -0.066225, -0.000100, 0.000000, -3.141593, 0.000000],accel_mss,speed_ms,0,0.000)
  movel(p[0.440613, -0.067066, -0.000100, 0.000000, -3.141593, 0.000000],accel_mss,speed_ms,0,0.000)
  movel(p[0.440672, -0.067504, -0.000100, 0.000000, -3.141593, 0.000000],accel_mss,speed_ms,0,0.000)
  movel(p[0.441118, -0.069267, -0.000100, 0.000000, -3.141593, 0.000000],accel_mss,speed_ms,0,0.001)
  movel(p[0.441698, -0.070864, -0.000100, 0.000000, -3.141593, 0.000000],accel_mss,speed_ms,0,0.001)
  movel(p[0.442378, -0.072220, -0.000100, 0.000000, -3.141593, 0.000000],accel_mss,speed_ms,0,0.001)
  movel(p[0.443124, -0.073245, -0.000100, 0.000000, 3.141593, 0.000000],accel_mss,speed_ms,0,0.001)
  movel(p[0.443383, -0.073542, -0.000100, 0.000000, -3.141593, 0.000000],accel_mss,speed_ms,0,0.000)
  movel(p[0.443602, -0.073812, -0.000100, 0.000000, 3.141593, 0.000000],accel_mss,speed_ms,0,0.000)
  movel(p[0.443776, -0.074042, -0.000100, 0.000000, -3.141593, 0.000000],accel_mss,speed_ms,0,0.000)
  movel(p[0.443861, -0.074283, -0.000100, 0.000000, -3.141593, 0.000000],accel_mss,speed_ms,0,0.000)
  movel(p[0.444135, -0.074587, -0.000100, 0.000000, 3.141593, 0.000000],accel_mss,speed_ms,0,0.000)
  movel(p[0.444432, -0.074868, -0.000100, 0.000000, -3.141593, 0.000000],accel_mss,speed_ms,0,0.000)
  movel(p[0.444594, -0.074929, -0.000100, 0.000000, -3.141593, 0.000000],accel_mss,speed_ms,0,0.000)
  movel(p[0.444942, -0.075141, -0.000100, 0.000000, -3.141593, 0.000000],accel_mss,speed_ms,0,0.000)
  movel(p[0.445246, -0.075374, -0.000100, 0.000000, -3.141593, 0.000000],accel_mss,speed_ms,0,0.000)
  movel(p[0.445580, -0.075651, -0.000100, 0.000000, -3.141593, 0.000000],accel_mss,speed_ms,0,0.000)
  movel(p[0.445948, -0.075947, -0.000100, 0.000000, -3.141593, 0.000000],accel_mss,speed_ms,0,0.000)
  movel(p[0.446354, -0.076238, -0.000100, 0.000000, -3.141593, 0.000000],accel_mss,speed_ms,0,0.000)
  movel(p[0.446737, -0.076484, -0.000100, 0.000000, -3.141593, 0.000000],accel_mss,speed_ms,0,0.000)
  movel(p[0.447026, -0.076633, -0.000100, 0.000000, -3.141593, 0.000000],accel_mss,speed_ms,0,0.000)
  movel(p[0.447275, -0.076743, -0.000100, 0.000000, -3.141593, 0.000000],accel_mss,speed_ms,0,0.000)
  movel(p[0.447526, -0.076859, -0.000100, 0.000000, -3.141593, 0.000000],accel_mss,speed_ms,0,0.000)
  movel(p[0.447748, -0.076964, -0.000100, 0.000000, -3.141593, 0.000000],accel_mss,speed_ms,0,0.000)
  movel(p[0.447888, -0.077036, -0.000100, 0.000000, -3.141593, 0.000000],accel_mss,speed_ms,0,0.000)
  movel(p[0.448338, -0.077274, -0.000100, 0.000000, -3.141593, 0.000000],accel_mss,speed_ms,0,0.000)
  movel(p[0.448678, -0.077438, -0.000100, 0.000000, -3.141593, 0.000000],accel_mss,speed_ms,0,0.000)
  movel(p[0.449060, -0.077598, -0.000100, 0.000000, -3.141593, 0.000000],accel_mss,speed_ms,0,0.000)
  movel(p[0.449672, -0.077836, -0.000100, 0.000000, 3.141593, 0.000000],accel_mss,speed_ms,0,0.000)
  movel(p[0.451635, -0.078440, -0.000100, 0.000000, -3.141593, 0.000000],accel_mss,speed_ms,0,0.001)
  movel(p[0.453365, -0.078663, -0.000100, 0.000000, -3.141593, 0.000000],accel_mss,speed_ms,0,0.001)
  movel(p[0.455170, -0.078524, -0.000100, 0.000000, -3.141593, 0.000000],accel_mss,speed_ms,0,0.001)
  movel(p[0.457378, -0.078012, -0.000100, 0.000000, -3.141593, 0.000000],accel_mss,speed_ms,0,0.001)
  movel(p[0.458203, -0.077753, -0.000100, 0.000000, -3.141593, 0.000000],accel_mss,speed_ms,0,0.000)
  movel(p[0.458842, -0.077496, -0.000100, 0.000000, -3.141593, 0.000000],accel_mss,speed_ms,0,0.000)
  movel(p[0.459469, -0.077170, -0.000100, 0.000000, -3.141593, 0.000000],accel_mss,speed_ms,0,0.000)
  movel(p[0.460260, -0.076686, -0.000100, 0.000000, -3.141593, 0.000000],accel_mss,speed_ms,0,0.000)
  movel(p[0.460513, -0.076530, -0.000100, 0.000000, -3.141593, 0.000000],accel_mss,speed_ms,0,0.000)
  movel(p[0.460749, -0.076399, -0.000100, 0.000000, -3.141593, 0.000000],accel_mss,speed_ms,0,0.000)
  movel(p[0.460949, -0.076298, -0.000100, 0.000000, -3.141593, 0.000000],accel_mss,speed_ms,0,0.000)
  movel(p[0.461285, -0.076177, -0.000100, 0.000000, -3.141593, 0.000000],accel_mss,speed_ms,0,0.000)
  movel(p[0.462184, -0.075296, -0.000100, 0.000000, -3.141593, 0.000000],accel_mss,speed_ms,0,0.001)
  movel(p[0.463027, -0.074426, -0.000100, 0.000000, -3.141593, 0.000000],accel_mss,speed_ms,0,0.000)
  movel(p[0.463297, -0.074016, -0.000100, 0.000000, 3.141593, 0.000000],accel_mss,speed_ms,0,0.000)
  movel(p[0.463379, -0.073846, -0.000100, 0.000000, 3.141593, 0.000000],accel_mss,speed_ms,0,0.000)
  movel(p[0.463496, -0.073628, -0.000100, 0.000000, -3.141593, 0.000000],accel_mss,speed_ms,0,0.000)
  movel(p[0.463626, -0.073403, -0.000100, 0.000000, -3.141593, 0.000000],accel_mss,speed_ms,0,0.000)
  movel(p[0.463751, -0.073204, -0.000100, 0.000000, -3.141593, 0.000000],accel_mss,speed_ms,0,0.000)
  movel(p[0.463872, -0.073015, -0.000100, 0.000000, -3.141593, 0.000000],accel_mss,speed_ms,0,0.000)
  movel(p[0.463991, -0.072820, -0.000100, 0.000000, -3.141593, 0.000000],accel_mss,speed_ms,0,0.000)
  movel(p[0.464091, -0.072645, -0.000100, 0.000000, -3.141593, 0.000000],accel_mss,speed_ms,0,0.000)
  movel(p[0.464150, -0.072529, -0.000100, 0.000000, -3.141593, 0.000000],accel_mss,speed_ms,0,0.000)
  movel(p[0.464211, -0.072413, -0.000100, 0.000000, 3.141593, 0.000000],accel_mss,speed_ms,0,0.000)
  movel(p[0.464318, -0.072238, -0.000100, 0.000000, -3.141593, 0.000000],accel_mss,speed_ms,0,0.000)
  movel(p[0.464445, -0.072043, -0.000100, 0.000000, -3.141593, 0.000000],accel_mss,speed_ms,0,0.000)
  movel(p[0.464576, -0.071854, -0.000100, 0.000000, -3.141593, 0.000000],accel_mss,speed_ms,0,0.000)
  movel(p[0.464819, -0.071468, -0.000100, 0.000000, -3.141593, 0.000000],accel_mss,speed_ms,0,0.000)
  movel(p[0.465165, -0.070810, -0.000100, 0.000000, -3.141593, 0.000000],accel_mss,speed_ms,0,0.000)
  movel(p[0.465641, -0.069844, -0.000100, 0.000000, -3.141593, 0.000000],accel_mss,speed_ms,0,0.000)
  movel(p[0.466342, -0.068367, -0.000100, 0.000000, -3.141593, 0.000000],accel_mss,speed_ms,0,0.001)
  movel(p[0.466486, -0.067832, -0.000100, 0.000000, -3.141593, 0.000000],accel_mss,speed_ms,0,0.000)
  movel(p[0.466501, -0.067062, -0.000100, 0.000000, 3.141593, 0.000000],accel_mss,speed_ms,0,0.000)
  movel(p[0.466411, -0.066307, -0.000100, 0.000000, -3.141593, 0.000000],accel_mss,speed_ms,0,0.000)
  movel(p[0.466215, -0.065828, -0.000100, 0.000000, -3.141593, 0.000000],accel_mss,speed_ms,0,0.000)
  movel(p[0.466094, -0.065644, -0.000100, 0.000000, -3.141593, 0.000000],accel_mss,speed_ms,0,0.000)
  movel(p[0.465968, -0.065441, -0.000100, 0.000000, 3.141593, 0.000000],accel_mss,speed_ms,0,0.000)
  movel(p[0.465854, -0.065250, -0.000100, 0.000000, -3.141593, 0.000000],accel_mss,speed_ms,0,0.000)
  movel(p[0.465774, -0.065107, -0.000100, 0.000000, -3.141593, 0.000000],accel_mss,speed_ms,0,0.000)
  movel(p[0.465693, -0.064982, -0.000100, 0.000000, -3.141593, 0.000000],accel_mss,speed_ms,0,0.000)
  movel(p[0.465576, -0.064852, -0.000100, 0.000000, -3.141593, 0.000000],accel_mss,speed_ms,0,0.000)
  movel(p[0.465443, -0.064737, -0.000100, 0.000000, -3.141593, 0.000000],accel_mss,speed_ms,0,0.000)
  movel(p[0.465315, -0.064657, -0.000100, 0.000000, 3.141593, 0.000000],accel_mss,speed_ms,0,0.000)
  movel(p[0.465156, -0.064565, -0.000100, 0.000000, -3.141593, 0.000000],accel_mss,speed_ms,0,0.000)
  movel(p[0.464906, -0.064395, -0.000100, 0.000000, -3.141593, 0.000000],accel_mss,speed_ms,0,0.000)
  movel(p[0.464626, -0.064191, -0.000100, 0.000000, 3.141593, 0.000000],accel_mss,speed_ms,0,0.000)
  movel(p[0.464351, -0.063979, -0.000100, 0.000000, -3.141593, 0.000000],accel_mss,speed_ms,0,0.000)
  movel(p[0.463895, -0.063628, -0.000100, 0.000000, -3.141593, 0.000000],accel_mss,speed_ms,0,0.000)
  movel(p[0.463517, -0.063362, -0.000100, 0.000000, -3.141593, 0.000000],accel_mss,speed_ms,0,0.000)
  movel(p[0.463179, -0.063155, -0.000100, 0.000000, -3.141593, 0.000000],accel_mss,speed_ms,0,0.000)
  movel(p[0.462851, -0.062988, -0.000100, 0.000000, -3.141593, 0.000000],accel_mss,speed_ms,0,0.000)
  movel(p[0.461472, -0.062388, -0.000100, 0.000000, -3.141593, 0.000000],accel_mss,speed_ms,0,0.001)
  movel(p[0.460432, -0.062010, -0.000100, 0.000000, -3.141593, 0.000000],accel_mss,speed_ms,0,0.000)
  movel(p[0.459592, -0.061798, -0.000100, 0.000000, 3.141593, 0.000000],accel_mss,speed_ms,0,0.000)
  movel(p[0.458856, -0.061729, -0.000100, 0.000000, 3.141593, 0.000000],accel_mss,speed_ms,0,0.000)
  movel(p[0.458180, -0.061784, -0.000100, 0.000000, -3.141593, 0.000000],accel_mss,speed_ms,0,0.000)
  movel(p[0.457371, -0.061955, -0.000100, 0.000000, -3.141593, 0.000000],accel_mss,speed_ms,0,0.000)
  movel(p[0.456628, -0.062179, -0.000100, 0.000000, -3.141593, 0.000000],accel_mss,speed_ms,0,0.000)
  movel(p[0.456253, -0.062402, -0.000100, 0.000000, -3.141593, 0.000000],accel_mss,speed_ms,0,0.000)
  movel(p[0.456146, -0.062489, -0.000100, 0.000000, -3.141593, 0.000000],accel_mss,speed_ms,0,0.000)
  movel(p[0.456033, -0.062562, -0.000100, 0.000000, -3.141593, 0.000000],accel_mss,speed_ms,0,0.000)
  movel(p[0.455930, -0.062614, -0.000100, 0.000000, -3.141593, 0.000000],accel_mss,speed_ms,0,0.000)
  movel(p[0.455652, -0.062712, -0.000100, 0.000000, -3.141593, 0.000000],accel_mss,speed_ms,0,0.000)
  movel(p[0.454992, -0.063367, -0.000100, 0.000000, -3.141593, 0.000000],accel_mss,speed_ms,0,0.000)
  movel(p[0.454375, -0.064022, -0.000100, 0.000000, -3.141593, 0.000000],accel_mss,speed_ms,0,0.000)
  movel(p[0.454064, -0.064450, -0.000100, 0.000000, -3.141593, 0.000000],accel_mss,speed_ms,0,0.000)
  movel(p[0.453631, -0.065275, -0.000100, 0.000000, 3.141593, 0.000000],accel_mss,speed_ms,0,0.000)
  movel(p[0.453438, -0.065876, -0.000100, 0.000000, 3.141593, 0.000000],accel_mss,speed_ms,0,0.000)
  movel(p[0.453445, -0.066359, -0.000100, 0.000000, -3.141593, 0.000000],accel_mss,speed_ms,0,0.000)
  movel(p[0.453635, -0.066796, -0.000100, 0.000000, -3.141593, 0.000000],accel_mss,speed_ms,0,0.000)
  movel(p[0.454260, -0.067319, -0.000100, 0.000000, -3.141593, 0.000000],accel_mss,speed_ms,0,0.000)
  movel(p[0.455269, -0.067637, -0.000100, 0.000000, -3.141593, 0.000000],accel_mss,speed_ms,0,0.000)
  movel(p[0.456363, -0.067699, -0.000100, 0.000000, -3.141593, 0.000000],accel_mss,speed_ms,0,0.000)
  movel(p[0.457253, -0.067453, -0.000100, 0.000000, -3.141593, 0.000000],accel_mss,speed_ms,0,0.000)
  movel(p[0.457514, -0.067301, -0.000100, 0.000000, -3.141593, 0.000000],accel_mss,speed_ms,0,0.000)
  movel(p[0.457796, -0.067100, -0.000100, 0.000000, -3.141593, 0.000000],accel_mss,speed_ms,0,0.000)
  movel(p[0.458054, -0.066885, -0.000100, 0.000000, -3.141593, 0.000000],accel_mss,speed_ms,0,0.000)
  movel(p[0.458244, -0.066689, -0.000100, 0.000000, -3.141593, 0.000000],accel_mss,speed_ms,0,0.000)
  movel(p[0.458504, -0.066316, -0.000100, 0.000000, -3.141593, 0.000000],accel_mss,speed_ms,0,0.000)
  movel(p[0.458746, -0.065833, -0.000100, 0.000000, -3.141593, 0.000000],accel_mss,speed_ms,0,0.000)
  movel(p[0.458921, -0.065365, -0.000100, 0.000000, -3.141593, 0.000000],accel_mss,speed_ms,0,0.000)
  movel(p[0.458939, -0.065084, -0.000100, 0.000000, -3.141593, 0.000000],accel_mss,speed_ms,0,0.000)
  movel(p[0.458904, -0.064805, -0.000100, 0.000000, -3.141593, 0.000000],accel_mss,speed_ms,0,0.000)
  movel(p[0.458955, -0.064705, -0.000100, 0.000000, -3.141593, 0.000000],accel_mss,speed_ms,0,0.000)
  movel(p[0.459177, -0.064934, -0.000100, 0.000000, -3.141593, 0.000000],accel_mss,speed_ms,0,0.000)
  movel(p[0.459385, -0.066013, -0.000100, 0.000000, -3.141593, 0.000000],accel_mss,speed_ms,0,0.000)
  movel(p[0.459009, -0.067183, -0.000100, 0.000000, -3.141593, 0.000000],accel_mss,speed_ms,0,0.000)
  movel(p[0.458131, -0.068200, -0.000100, 0.000000, -3.141593, 0.000000],accel_mss,speed_ms,0,0.001)
  movel(p[0.456926, -0.068839, -0.000100, 0.000000, -3.141593, 0.000000],accel_mss,speed_ms,0,0.001)
  movel(p[0.455025, -0.069127, -0.000100, 0.000000, 3.141593, 0.000000],accel_mss,speed_ms,0,0.001)
  movel(p[0.453288, -0.068774, -0.000100, 0.000000, -3.141593, 0.000000],accel_mss,speed_ms,0,0.001)
  movel(p[0.451988, -0.067843, -0.000100, 0.000000, 3.141593, 0.000000],accel_mss,speed_ms,0,0.001)
  movel(p[0.451307, -0.066484, -0.000100, 0.000000, -3.141593, 0.000000],accel_mss,speed_ms,0,0.001)
  movel(p[0.451251, -0.065080, -0.000100, 0.000000, 3.141593, 0.000000],accel_mss,speed_ms,0,0.001)
  movel(p[0.451635, -0.063587, -0.000100, 0.000000, 3.141593, 0.000000],accel_mss,speed_ms,0,0.001)
  movel(p[0.452430, -0.062102, -0.000100, 0.000000, -3.141593, 0.000000],accel_mss,speed_ms,0,0.001)
  movel(p[0.453590, -0.060723, -0.000100, 0.000000, -3.141593, 0.000000],accel_mss,speed_ms,0,0.001)
  movel(p[0.454308, -0.060048, -0.000100, 0.000000, -3.141593, 0.000000],accel_mss,speed_ms,0,0.000)
  movel(p[0.454914, -0.059554, -0.000100, 0.000000, -3.141593, 0.000000],accel_mss,speed_ms,0,0.000)
  movel(p[0.455484, -0.059180, -0.000100, 0.000000, 3.141593, 0.000000],accel_mss,speed_ms,0,0.000)
  movel(p[0.456088, -0.058875, -0.000100, 0.000000, -3.141593, 0.000000],accel_mss,speed_ms,0,0.000)
  movel(p[0.456256, -0.058791, -0.000100, 0.000000, -3.141593, 0.000000],accel_mss,speed_ms,0,0.000)
  movel(p[0.456332, -0.058715, -0.000100, 0.000000, -3.141593, 0.000000],accel_mss,speed_ms,0,0.000)
  movel(p[0.456280, -0.058548, -0.000100, 0.000000, -3.141593, 0.000000],accel_mss,speed_ms,0,0.000)
  movel(p[0.456262, -0.058395, -0.000100, 0.000000, -3.141593, 0.000000],accel_mss,speed_ms,0,0.000)
  movel(p[0.456509, -0.058042, -0.000100, 0.000000, -3.141593, 0.000000],accel_mss,speed_ms,0,0.000)
  movel(p[0.456958, -0.057519, -0.000100, 0.000000, -3.141593, 0.000000],accel_mss,speed_ms,0,0.000)
  movel(p[0.457747, -0.056688, -0.000100, 0.000000, -3.141593, 0.000000],accel_mss,speed_ms,0,0.000)
  movel(p[0.458670, -0.055686, -0.000100, 0.000000, 3.141593, 0.000000],accel_mss,speed_ms,0,0.001)
  movel(p[0.459366, -0.054814, -0.000100, 0.000000, -3.141593, 0.000000],accel_mss,speed_ms,0,0.000)
  movel(p[0.459845, -0.054071, -0.000100, 0.000000, -3.141593, 0.000000],accel_mss,speed_ms,0,0.000)
  movel(p[0.460078, -0.053479, -0.000100, 0.000000, -3.141593, 0.000000],accel_mss,speed_ms,0,0.000)
  movel(p[0.460204, -0.053184, -0.000100, 0.000000, -3.141593, 0.000000],accel_mss,speed_ms,0,0.000)
  movel(p[0.460332, -0.052900, -0.000100, 0.000000, -3.141593, 0.000000],accel_mss,speed_ms,0,0.000)
  movel(p[0.460480, -0.052579, -0.000100, 0.000000, -3.141593, 0.000000],accel_mss,speed_ms,0,0.000)
  movel(p[0.460854, -0.051737, -0.000100, 0.000000, -3.141593, 0.000000],accel_mss,speed_ms,0,0.000)
  movel(p[0.461074, -0.051129, -0.000100, 0.000000, -3.141593, 0.000000],accel_mss,speed_ms,0,0.000)
  movel(p[0.461176, -0.050686, -0.000100, 0.000000, -3.141593, 0.000000],accel_mss,speed_ms,0,0.000)
  movel(p[0.461146, -0.050402, -0.000100, 0.000000, -3.141593, 0.000000],accel_mss,speed_ms,0,0.000)
  movel(p[0.461078, -0.050253, -0.000100, 0.000000, -3.141593, 0.000000],accel_mss,speed_ms,0,0.000)
  movel(p[0.460941, -0.050241, -0.000100, 0.000000, -3.141593, 0.000000],accel_mss,speed_ms,0,0.000)
  movel(p[0.460773, -0.050384, -0.000100, 0.000000, -3.141593, 0.000000],accel_mss,speed_ms,0,0.000)
  movel(p[0.460659, -0.050477, -0.000100, 0.000000, -3.141593, 0.000000],accel_mss,speed_ms,0,0.000)
  movel(p[0.460539, -0.050557, -0.000100, 0.000000, 3.141593, 0.000000],accel_mss,speed_ms,0,0.000)
  movel(p[0.460430, -0.050613, -0.000100, 0.000000, -3.141593, 0.000000],accel_mss,speed_ms,0,0.000)
  movel(p[0.460273, -0.050655, -0.000100, 0.000000, 3.141593, 0.000000],accel_mss,speed_ms,0,0.000)
  movel(p[0.460103, -0.050783, -0.000100, 0.000000, -3.141593, 0.000000],accel_mss,speed_ms,0,0.000)
  movel(p[0.459906, -0.050953, -0.000100, 0.000000, -3.141593, 0.000000],accel_mss,speed_ms,0,0.000)
  movel(p[0.459701, -0.051154, -0.000100, 0.000000, -3.141593, 0.000000],accel_mss,speed_ms,0,0.000)
  movel(p[0.459495, -0.051355, -0.000100, 0.000000, 3.141593, 0.000000],accel_mss,speed_ms,0,0.000)
  movel(p[0.459299, -0.051525, -0.000100, 0.000000, -3.141593, 0.000000],accel_mss,speed_ms,0,0.000)
  movel(p[0.459130, -0.051653, -0.000100, 0.000000, -3.141593, 0.000000],accel_mss,speed_ms,0,0.000)
  movel(p[0.458966, -0.051698, -0.000100, 0.000000, 3.141593, 0.000000],accel_mss,speed_ms,0,0.000)
  movel(p[0.458810, -0.051780, -0.000100, 0.000000, -3.141593, 0.000000],accel_mss,speed_ms,0,0.000)
  movel(p[0.458628, -0.051892, -0.000100, 0.000000, -3.141593, 0.000000],accel_mss,speed_ms,0,0.000)
  movel(p[0.458440, -0.052025, -0.000100, 0.000000, -3.141593, 0.000000],accel_mss,speed_ms,0,0.000)
  movel(p[0.458036, -0.052289, -0.000100, 0.000000, -3.141593, 0.000000],accel_mss,speed_ms,0,0.000)
  movel(p[0.457444, -0.052609, -0.000100, 0.000000, -3.141593, 0.000000],accel_mss,speed_ms,0,0.000)
  movel(p[0.456698, -0.052972, -0.000100, 0.000000, -3.141593, 0.000000],accel_mss,speed_ms,0,0.000)
  movel(p[0.455801, -0.053375, -0.000100, 0.000000, -3.141593, 0.000000],accel_mss,speed_ms,0,0.000)
  movel(p[0.455556, -0.053469, -0.000100, 0.000000, -3.141593, 0.000000],accel_mss,speed_ms,0,0.000)
  movel(p[0.455254, -0.053564, -0.000100, 0.000000, 3.141593, 0.000000],accel_mss,speed_ms,0,0.000)
  movel(p[0.454943, -0.053645, -0.000100, 0.000000, -3.141593, 0.000000],accel_mss,speed_ms,0,0.000)
  movel(p[0.454676, -0.053699, -0.000100, 0.000000, -3.141593, 0.000000],accel_mss,speed_ms,0,0.000)
  movel(p[0.454424, -0.053742, -0.000100, 0.000000, -3.141593, 0.000000],accel_mss,speed_ms,0,0.000)
  movel(p[0.454164, -0.053792, -0.000100, 0.000000, -3.141593, 0.000000],accel_mss,speed_ms,0,0.000)
  movel(p[0.453931, -0.053841, -0.000100, 0.000000, -3.141593, 0.000000],accel_mss,speed_ms,0,0.000)
  movel(p[0.453776, -0.053881, -0.000100, 0.000000, -3.141593, 0.000000],accel_mss,speed_ms,0,0.000)
  movel(p[0.453611, -0.053919, -0.000100, 0.000000, 3.141593, 0.000000],accel_mss,speed_ms,0,0.000)
  movel(p[0.453619, -0.053815, -0.000100, 0.000000, 3.141593, 0.000000],accel_mss,speed_ms,0,0.000)
  movel(p[0.453839, -0.053573, -0.000100, 0.000000, -3.141593, 0.000000],accel_mss,speed_ms,0,0.000)
  movel(p[0.453990, -0.053422, -0.000100, 0.000000, -3.141593, 0.000000],accel_mss,speed_ms,0,0.000)
  movel(p[0.454143, -0.053294, -0.000100, 0.000000, -3.141593, 0.000000],accel_mss,speed_ms,0,0.000)
  movel(p[0.454280, -0.053201, -0.000100, 0.000000, -3.141593, 0.000000],accel_mss,speed_ms,0,0.000)
  movel(p[0.454467, -0.053141, -0.000100, 0.000000, -3.141593, 0.000000],accel_mss,speed_ms,0,0.000)
  movel(p[0.454831, -0.052851, -0.000100, 0.000000, -3.141593, 0.000000],accel_mss,speed_ms,0,0.000)
  movel(p[0.455254, -0.052494, -0.000100, 0.000000, -3.141593, 0.000000],accel_mss,speed_ms,0,0.000)
  movel(p[0.455726, -0.052070, -0.000100, 0.000000, -3.141593, 0.000000],accel_mss,speed_ms,0,0.000)
  movel(p[0.456326, -0.051518, -0.000100, 0.000000, -3.141593, 0.000000],accel_mss,speed_ms,0,0.000)
  movel(p[0.456926, -0.050965, -0.000100, 0.000000, -3.141593, 0.000000],accel_mss,speed_ms,0,0.000)
  movel(p[0.456738, -0.050804, -0.000100, 0.000000, -3.141593, 0.000000],accel_mss,speed_ms,0,0.000)
  movel(p[0.456551, -0.050642, -0.000100, 0.000000, -3.141593, 0.000000],accel_mss,speed_ms,0,0.000)
  movel(p[0.456382, -0.050508, -0.000100, 0.000000, -3.141593, 0.000000],accel_mss,speed_ms,0,0.000)
  movel(p[0.456187, -0.050372, -0.000100, 0.000000, -3.141593, 0.000000],accel_mss,speed_ms,0,0.000)
  movel(p[0.455994, -0.050254, -0.000100, 0.000000, -3.141593, 0.000000],accel_mss,speed_ms,0,0.000)
  movel(p[0.455838, -0.050177, -0.000100, 0.000000, 3.141593, 0.000000],accel_mss,speed_ms,0,0.000)
  movel(p[0.455624, -0.049995, -0.000100, 0.000000, 3.141593, 0.000000],accel_mss,speed_ms,0,0.000)
  movel(p[0.455507, -0.049685, -0.000100, 0.000000, -3.141593, 0.000000],accel_mss,speed_ms,0,0.000)
  movel(p[0.455509, -0.049322, -0.000100, 0.000000, -3.141593, 0.000000],accel_mss,speed_ms,0,0.000)
  movel(p[0.455638, -0.048995, -0.000100, 0.000000, -3.141593, 0.000000],accel_mss,speed_ms,0,0.000)
  movel(p[0.455763, -0.048888, -0.000100, 0.000000, 3.141593, 0.000000],accel_mss,speed_ms,0,0.000)
  movel(p[0.455918, -0.048877, -0.000100, 0.000000, 3.141593, 0.000000],accel_mss,speed_ms,0,0.000)
  movel(p[0.456158, -0.048983, -0.000100, 0.000000, -3.141593, 0.000000],accel_mss,speed_ms,0,0.000)
  movel(p[0.456626, -0.049278, -0.000100, 0.000000, 3.141593, 0.000000],accel_mss,speed_ms,0,0.000)
  movel(p[0.456820, -0.049403, -0.000100, 0.000000, -3.141593, 0.000000],accel_mss,speed_ms,0,0.000)
  movel(p[0.457032, -0.049532, -0.000100, 0.000000, -3.141593, 0.000000],accel_mss,speed_ms,0,0.000)
  movel(p[0.457229, -0.049648, -0.000100, 0.000000, -3.141593, 0.000000],accel_mss,speed_ms,0,0.000)
  movel(p[0.457376, -0.049726, -0.000100, 0.000000, -3.141593, 0.000000],accel_mss,speed_ms,0,0.000)
  movel(p[0.457509, -0.049798, -0.000100, 0.000000, -3.141593, 0.000000],accel_mss,speed_ms,0,0.000)
  movel(p[0.457663, -0.049888, -0.000100, 0.000000, -3.141593, 0.000000],accel_mss,speed_ms,0,0.000)
  movel(p[0.457813, -0.049981, -0.000100, 0.000000, -3.141593, 0.000000],accel_mss,speed_ms,0,0.000)
  movel(p[0.457933, -0.050062, -0.000100, 0.000000, 3.141593, 0.000000],accel_mss,speed_ms,0,0.000)
  movel(p[0.458085, -0.050138, -0.000100, 0.000000, 3.141593, 0.000000],accel_mss,speed_ms,0,0.000)
  movel(p[0.458220, -0.050138, -0.000100, 0.000000, -3.141593, 0.000000],accel_mss,speed_ms,0,0.000)
  movel(p[0.458374, -0.050057, -0.000100, 0.000000, -3.141593, 0.000000],accel_mss,speed_ms,0,0.000)
  movel(p[0.458608, -0.049856, -0.000100, 0.000000, -3.141593, 0.000000],accel_mss,speed_ms,0,0.000)
  movel(p[0.458781, -0.049703, -0.000100, 0.000000, -3.141593, 0.000000],accel_mss,speed_ms,0,0.000)
  movel(p[0.458954, -0.049564, -0.000100, 0.000000, -3.141593, 0.000000],accel_mss,speed_ms,0,0.000)
  movel(p[0.459108, -0.049455, -0.000100, 0.000000, -3.141593, 0.000000],accel_mss,speed_ms,0,0.000)
  movel(p[0.459201, -0.049410, -0.000100, 0.000000, -3.141593, 0.000000],accel_mss,speed_ms,0,0.000)
  movel(p[0.459315, -0.049350, -0.000100, 0.000000, -3.141593, 0.000000],accel_mss,speed_ms,0,0.000)
  movel(p[0.459714, -0.049032, -0.000100, 0.000000, 3.141593, 0.000000],accel_mss,speed_ms,0,0.000)
  movel(p[0.460181, -0.048647, -0.000100, 0.000000, -3.141593, 0.000000],accel_mss,speed_ms,0,0.000)
  movel(p[0.460701, -0.048201, -0.000100, 0.000000, -3.141593, 0.000000],accel_mss,speed_ms,0,0.000)
  movel(p[0.462085, -0.046990, -0.000100, 0.000000, -3.141593, 0.000000],accel_mss,speed_ms,0,0.001)
  movel(p[0.462714, -0.046416, -0.000100, 0.000000, -3.141593, 0.000000],accel_mss,speed_ms,0,0.000)
  movel(p[0.463064, -0.046063, -0.000100, 0.000000, -3.141593, 0.000000],accel_mss,speed_ms,0,0.000)
  movel(p[0.463140, -0.045885, -0.000100, 0.000000, -3.141593, 0.000000],accel_mss,speed_ms,0,0.000)
  movel(p[0.463215, -0.045710, -0.000100, 0.000000, -3.141593, 0.000000],accel_mss,speed_ms,0,0.000)
